(* IEC 61131-3 sources: STruCpp/libs/sources/plcopen-softmotion, 17 files *)

(* ---- opensml_axis.st ---- *)
(*
 * OpenSML_Axis — CiA 402 axis reference structure.
 *
 * Vendored from OpenSML (https://github.com/feecat/OpenSML), GPL-3.0.
 * Each field maps 1:1 onto a CiA 402 drive object exchanged over the
 * fieldbus (e.g. EtherCAT PDOs). Outputs (%Q) are written by the motion
 * blocks; inputs (%I) are read from the drive each scan.
 *)
TYPE OpenSML_Axis :
STRUCT
	(* Outputs -> drive *)
	ControlWord : UINT;                 (* 0x6040 *)
	Modes_of_operation : SINT;          (* 0x6060 *)
	Target_Position : DINT;             (* 0x607A *)
	Profile_Velocity : UDINT;           (* 0x6081 *)
	Target_Velocity : DINT;             (* 0x60FF *)
	Target_torque : INT;                (* 0x6071 *)
	(* Inputs <- drive *)
	StatusWord : UINT;                  (* 0x6041 *)
	Modes_of_operation_display : SINT;  (* 0x6061 *)
	Torque_Actual_Value : INT;          (* 0x6077 *)
	Position_Actual_Value : DINT;       (* 0x6064 *)
	Velocity_Actual_Value : DINT;       (* 0x606C *)
	Current_Actual_Value : INT;         (* 0x6078 *)
	Following_Error_Actual_Value : DINT;(* 0x60F4 *)
END_STRUCT
END_TYPE

(* ---- opensml_control.st ---- *)
(*
 * OpenSML_Control — aggregate axis command/status structure.
 * Vendored from OpenSML (https://github.com/feecat/OpenSML), GPL-3.0.
 *)
TYPE OpenSML_Control :
STRUCT
	xAxisEnable: BOOL;//Axis Hardware Enable
	xMoveEnable: BOOL;//Jog&Pos Movement Enable
	xHomeEnable: BOOL;//Home Function Enable
	xSimulation: BOOL;//Simulation Mode
	xEmergencyStop: BOOL:=TRUE;//Emergency Stop

	JogPos: BOOL;//Jog Positive
	JogNeg: BOOL;//Jog Negative
	JogVelocity: LREAL:=10;//Jog Velocity

	lrActualPosition: LREAL;//Actual Position Feedback

	lrFollowPosition: LREAL;//Follow Target Position, Can be set to new value at any time
	lrFollowVelocity: LREAL:=20;//Follow Move Velocity, Can be set to new value at any time
	xFollowEnable: BOOL;//Follow Move Enable

	xError: BOOL;//Error
	xBusy: BOOL;//Busy, Normal Working State
	xInPosition: BOOL;//In Position
	xEnabled: BOOL;//Axis Hardware Enabled
	xHomeDone: BOOL;//Axis Home Done

	MaxVelocity: LREAL:=100;//Max Velocity
	MaxAcceleration: LREAL:=1000;//Max Acceleration
	MaxJerk: LREAL:=10000;//Max Jerk
	CycleTime: LREAL:=0.001;//Task Cycle Time, 0.001 = 1ms
	Scale: LREAL:=16#1000;//Scale

	Axis:OpenSML_Axis;//Axis Reference
END_STRUCT
END_TYPE

(* ---- s7rtt_types.st ---- *)
(*
 * S7RTT motion-state / limits structures.
 * Vendored from S7RTT (https://github.com/feecat/S7RTT), Apache-2.0.
 * Converted from PLCopen XML. Single-axis 7-segment S-curve OTG.
 *)

TYPE ST_MotionLimits :
STRUCT
	fVelMax : LREAL;
	fAccMax : LREAL;
	fJerkMax : LREAL;
END_STRUCT
END_TYPE

TYPE ST_MotionState :
STRUCT
	fDuration : LREAL := 0.0;
	fPos : LREAL := 0.0;
	fVel : LREAL := 0.0;
	fAcc : LREAL := 0.0;
	fJerk : LREAL := 0.0;
END_STRUCT
END_TYPE

(* ---- sm3_axis_ref.st ---- *)
(*
 * AXIS_REF_SM3 — CODESYS SoftMotion-compatible axis reference.
 *
 * Application code declares an axis of this type (the EtherCAT drive's name),
 * passes it to MC_* blocks by VAR_IN_OUT, and reads/writes its fields
 * (fActPosition, nAxisState, …) — exactly as in CODESYS. It is a STRUCT (not an
 * FB): real CODESYS application code never calls axis methods (those are all
 * driver-internal). All positions/velocities are in technical (user) units;
 * the embedded `Drive` carries the raw CiA 402 PDO words in increments, and
 * SM_Drive_GenericDS402 bridges between them each scan.
 *)
TYPE AXIS_REF_SM3 :
STRUCT
	(* --- Command (written by MC_* blocks, in technical units) --- *)
	fSetPosition : LREAL;              (* commanded position [u] *)
	fSetVelocity : LREAL;              (* commanded velocity [u/s] *)
	fSetAcceleration : LREAL;          (* commanded acceleration [u/s2] *)
	fSetDeceleration : LREAL;          (* commanded deceleration [u/s2] *)
	fSetJerk : LREAL;                  (* commanded jerk [u/s3] *)
	bRegulatorOn : BOOL;               (* power-stage enable command *)
	bDriveStart : BOOL;                (* quick-stop release command *)
	byControllerMode : BYTE;           (* SMC_CONTROLLER_MODE as BYTE *)

	(* --- Feedback (updated by the drive bridge, in technical units) --- *)
	fActPosition : LREAL;              (* actual position [u] *)
	fActVelocity : LREAL;              (* actual velocity [u/s] *)
	fActTorque : LREAL;                (* actual torque *)
	nAxisState : SMC_AXIS_STATE;       (* PLCopen axis state *)
	bRegulatorRealState : BOOL;        (* real power-stage state *)
	bDriveStartRealState : BOOL;       (* real quick-stop-released state *)
	byRealControllerMode : BYTE;       (* actual controller mode *)

	(* --- Error / communication --- *)
	bError : BOOL;
	dwErrorID : DWORD;                 (* SMC_ERROR as DWORD *)
	bCommunication : BOOL;
	wCommunicationState : WORD;

	(* --- Scaling (increments <-> technical units) --- *)
	iRatioTechUnitsNum : DINT := 1;    (* CODESYS param 1052 *)
	dwRatioTechUnitsDenom : DWORD := 1;(* CODESYS param 1051 *)
	fScalefactor : LREAL := 1.0;       (* CODESYS param 1054 *)
	fIncPerUnit : LREAL := 1.0;        (* derived: increments per user unit *)

	(* --- Axis configuration --- *)
	fPositionPeriod : LREAL := 360.0;  (* modulo period [u] *)
	bModulo : BOOL;                    (* TRUE = rotary/modulo axis *)
	fSWLimitPositive : LREAL;
	fSWLimitNegative : LREAL;
	bSWLimitEnable : BOOL;
	fCycleTime : LREAL := 0.01;        (* task cycle [s], for OTG *)

	(* --- Raw CiA 402 interface (increments) bridged to the drive PDOs --- *)
	Drive : OpenSML_Axis;
END_STRUCT
END_TYPE

(* ---- sm3_enums.st ---- *)
(*
 * CODESYS SoftMotion (SM3) compatible enum types.
 *
 * Values follow CODESYS SM3_Basic / SM3_Error so that ported application code
 * comparing against these names/values behaves identically. This is the
 * single-axis CiA 402 subset (see docs/PLCOPEN_SOFTMOTION_ETHERCAT_PLAN.md).
 *)

(* PLCopen axis state (AXIS_REF_SM3.nAxisState) *)
TYPE SMC_AXIS_STATE : (
	power_off := 0,
	errorstop := 1,
	stopping := 2,
	standstill := 3,
	discrete_motion := 4,
	continuous_motion := 5,
	synchronized_motion := 6,
	homing := 7
); END_TYPE

(* Controller mode (AXIS_REF_SM3.byControllerMode / SMC_SetControllerMode) *)
TYPE SMC_CONTROLLER_MODE : (
	SMC_nocontrol := 0,
	SMC_torque := 1,
	SMC_velocity := 2,
	SMC_position := 3,
	SMC_current := 4
); END_TYPE

(* Movement direction for MC_MoveAbsolute / MC_MoveVelocity (modulo axes) *)
TYPE MC_DIRECTION : (
	mcd_negative := -1,
	mcd_current := 0,
	mcd_positive := 1,
	mcd_shortest := 2,
	mcd_fastest := 3
); END_TYPE

(* Buffering behaviour relative to a preceding motion command *)
TYPE MC_BUFFER_MODE : (
	mcbm_aborting := 0,
	mcbm_buffered := 1,
	mcbm_blending_low := 2,
	mcbm_blending_previous := 3,
	mcbm_blending_next := 4,
	mcbm_blending_high := 5
); END_TYPE

(* Homing mode (subset — the CiA 402 relevant ones) *)
TYPE SMC_HOMING_MODE : (
	smc_hm_direct := 0,
	smc_hm_limit_switch := 1,
	smc_hm_reference_pulse := 2,
	smc_hm_drive_internal := 35
); END_TYPE

(*
 * Error identifier (MC_*.ErrorID). Single-axis CiA 402 subset of CODESYS
 * SMC_ERROR (the 0..~500 drive-interface / limits / controller-mode /
 * FB-input band). Values match CODESYS where documented.
 *)
TYPE SMC_ERROR : (
	SMC_NO_ERROR := 0,
	SMC_DI_GENERAL_COMMUNICATION_ERROR := 1,
	SMC_DI_AXIS_ERROR := 2,
	SMC_DI_SWLIMITS_EXCEEDED := 10,
	SMC_DI_HWLIMITS_EXCEEDED := 11,
	SMC_DI_HALT_OR_QUICKSTOP_NOT_SUPPORTED := 12,
	SMC_DI_VOLTAGE_DISABLED := 13,
	SMC_DI_FIELDBUS_LOST_SYNCRONITY := 14,
	SMC_DI_COMMUNICATION_INTERRUPTED := 15,
	SMC_REGULATOR_OR_START_NOT_SET := 20,
	SMC_WRONG_CONTROLLER_MODE := 21,
	SMC_FB_WASNT_CALLED_DURING_MOTION := 22,
	SMC_AXIS_IS_NO_AXIS_REF := 23,
	SMC_AXIS_REF_CHANGED_DURING_OPERATION := 24,
	SMC_FB_ACTIVE_AXIS_DISABLED := 25,
	SMC_AXIS_NOT_READY_FOR_MOTION := 26,
	SMC_NicNyet_ERROR := 30,
	SMC_MA_INVALID_ACCDEC_VALUES := 110,
	SMC_MA_INVALID_DIRECTION := 111,
	SMC_MV_INVALID_VELACC_VALUES := 120,
	SMC_MV_DIRECTION_NOT_APPLICABLE := 121,
	SMC_H_AXIS_WASNT_STANDING_STILL := 130,
	SMC_H_AXIS_DIDNT_START_HOMING := 131,
	SMC_H_HOMING_TIMEOUT := 132,
	SMC_R_NO_ERROR_TO_RESET := 140,
	SMC_R_DRIVE_DOESNT_ANSWER := 141,
	SMC_STOP_ERROR_DURING_STOP := 150,
	SMC_3SH_INVALID_VELACC_VALUES := 160
); END_TYPE

(* ---- s7rtt_functions.st ---- *)
(*
 * S7RTT trajectory helper functions (AtTime / BuildProfile / CalcTrajDist).
 * Vendored from S7RTT (https://github.com/feecat/S7RTT), Apache-2.0.
 * Converted from PLCopen XML. Single-axis 7-segment S-curve OTG.
 *)

FUNCTION FC_S7RTT_AtTime : ST_MotionState
VAR_INPUT
	Trajectory : ARRAY[1..32] OF ST_MotionState;
	SegCount : INT;
	ElapsedTime : LREAL;
END_VAR
VAR
	i : INT;
	t_rem : LREAL;
	t : LREAL;
	j : LREAL;
	p0 : LREAL;
	v0 : LREAL;
	a0 : LREAL;
	last_idx : INT;
END_VAR

IF SegCount <= 0 THEN
    // No trajectory, return first state
    FC_S7RTT_AtTime.fPos := Trajectory[1].fPos; FC_S7RTT_AtTime.fVel := 0.0; FC_S7RTT_AtTime.fAcc := 0.0;
    RETURN;
END_IF;

IF ElapsedTime <= 0.0 THEN
     // Return Initial State from First Segment
     FC_S7RTT_AtTime := Trajectory[1];
     FC_S7RTT_AtTime.fDuration := 0.0;
     FC_S7RTT_AtTime.fJerk := 0.0;
     RETURN;
END_IF;

t_rem := ElapsedTime;

FOR i := 1 TO SegCount DO
	IF t_rem <= Trajectory[i].fDuration THEN
		t := t_rem;
		j := Trajectory[i].fJerk;
		// Use pre-calculated state at segment start
		p0 := Trajectory[i].fPos;
		v0 := Trajectory[i].fVel;
		a0 := Trajectory[i].fAcc;

		FC_S7RTT_AtTime.fPos := p0 + v0 * t + 0.5 * a0 * t*t + (1.0/6.0) * j * t*t*t;
		FC_S7RTT_AtTime.fVel := v0 + a0 * t + 0.5 * j * t*t;
		FC_S7RTT_AtTime.fAcc := a0 + j * t;
		FC_S7RTT_AtTime.fJerk := j;
		FC_S7RTT_AtTime.fDuration := 0.0;
		RETURN;
	ELSE
		t_rem := t_rem - Trajectory[i].fDuration;
	END_IF;
END_FOR;

// Time is beyond end of trajectory
// Calculate Final State of last segment
last_idx := SegCount;
t := Trajectory[last_idx].fDuration;
j := Trajectory[last_idx].fJerk;
p0 := Trajectory[last_idx].fPos;
v0 := Trajectory[last_idx].fVel;
a0 := Trajectory[last_idx].fAcc;

p0 := p0 + v0 * t + 0.5 * a0 * t*t + (1.0/6.0) * j * t*t*t;
v0 := v0 + a0 * t + 0.5 * j * t*t;

// Hold Final Position (assuming v=target, a=0 at end)
// Linear projection if Velocity is non-zero
FC_S7RTT_AtTime.fPos := p0 + v0 * t_rem;
FC_S7RTT_AtTime.fVel := v0;
FC_S7RTT_AtTime.fAcc := 0.0;
FC_S7RTT_AtTime.fJerk := 0.0;
FC_S7RTT_AtTime.fDuration := 0.0;
END_FUNCTION

FUNCTION FC_S7RTT_BuildProfile : INT
VAR_INPUT
	in_v_start : LREAL;
	in_a_start : LREAL;
	in_v_target : LREAL;
	in_a_max : LREAL;
	in_j_max : LREAL;
END_VAR
VAR_IN_OUT
	out_time : ARRAY[1..5] OF LREAL;
	out_jerk : ARRAY[1..5] OF LREAL;
END_VAR
VAR
	acc_clamped : LREAL;
	t_to_zero : LREAL;
	j_restore : LREAL;
	v_min_feasible : LREAL;
	direction : LREAL;
	v0_mod : LREAL;
	a0_mod : LREAL;
	v1_mod : LREAL;
	t1_max : LREAL;
	t3_max : LREAL;
	dv_inflection : LREAL;
	dv_req : LREAL;
	dv_missing : LREAL;
	term : LREAL;
	a_peak : LREAL;
	t1 : LREAL;
	t2 : LREAL;
	t3 : LREAL;
	cnt : INT;
	EPS : LREAL := 1E-10;
END_VAR

cnt := 0;

// 1. Clamp initial acceleration to limits
acc_clamped := in_a_start;
IF acc_clamped > in_a_max THEN acc_clamped := in_a_max; END_IF;
IF acc_clamped < -in_a_max THEN acc_clamped := -in_a_max; END_IF;

// 2. Check feasibility (can we stop?)
t_to_zero := ABS(acc_clamped) / in_j_max;
IF ABS(acc_clamped) > EPS THEN
    IF acc_clamped > 0.0 THEN j_restore := -in_j_max; ELSE j_restore := in_j_max; END_IF;
ELSE
    j_restore := 0.0;
END_IF;

v_min_feasible := in_v_start + acc_clamped * t_to_zero + 0.5 * j_restore * t_to_zero * t_to_zero;

// 3. Determine direction
direction := 1.0;
IF in_v_target < v_min_feasible - EPS THEN
    direction := -1.0;
END_IF;

// 4. Normalize to positive quadrant
v0_mod := in_v_start * direction;
a0_mod := acc_clamped * direction;
v1_mod := in_v_target * direction;

t1_max := (in_a_max - a0_mod) / in_j_max;
IF t1_max < 0.0 THEN t1_max := 0.0; END_IF;

t3_max := in_a_max / in_j_max;

// Velocity change at inflection (max accel reached)
dv_inflection := (a0_mod * t1_max + 0.5 * in_j_max * t1_max * t1_max) +
                 (in_a_max * t3_max - 0.5 * in_j_max * t3_max * t3_max);

dv_req := v1_mod - v0_mod;

// 5. Calculate profile times
IF dv_req > dv_inflection THEN
    // Trapezoidal (Constant Acceleration Phase)
    dv_missing := dv_req - dv_inflection;
    t2 := dv_missing / in_a_max;
    t1 := t1_max;
    t3 := t3_max;
ELSE
    // Triangular (No Constant Acceleration)
    term := in_j_max * dv_req + 0.5 * a0_mod * a0_mod;
    IF term < 0.0 THEN term := 0.0; END_IF;
    a_peak := SQRT(term);

    t1 := (a_peak - a0_mod) / in_j_max;
    IF t1 < 0.0 THEN t1 := 0.0; END_IF;

    t3 := a_peak / in_j_max;
    IF t3 < 0.0 THEN t3 := 0.0; END_IF;

    t2 := 0.0;
END_IF;

// 6. Output Segments
IF t1 > EPS THEN
    cnt := cnt + 1; out_time[cnt] := t1; out_jerk[cnt] := direction * in_j_max;
END_IF;
IF t2 > EPS THEN
    cnt := cnt + 1; out_time[cnt] := t2; out_jerk[cnt] := 0.0;
END_IF;
IF t3 > EPS THEN
    cnt := cnt + 1; out_time[cnt] := t3; out_jerk[cnt] := -direction * in_j_max;
END_IF;

FC_S7RTT_BuildProfile := cnt;
END_FUNCTION

FUNCTION FC_S7RTT_CalcTrajDist : LREAL
VAR_INPUT
	v_peak : LREAL;
	start_v : LREAL;
	start_a : LREAL;
	target_v : LREAL;
	a_max : LREAL;
	j_max : LREAL;
END_VAR
VAR
	t_buf : ARRAY[1..5] OF LREAL;
	j_buf : ARRAY[1..5] OF LREAL;
	cnt : INT;
	i : INT;
	v_curr : LREAL;
	a_curr : LREAL;
	dist_total : LREAL;
	t_seg : LREAL;
	j_seg : LREAL;
END_VAR

dist_total := 0.0;
v_curr := start_v;
a_curr := start_a;

// Phase 1: Start -> Peak Velocity
cnt := FC_S7RTT_BuildProfile(v_curr, a_curr, v_peak, a_max, j_max, t_buf, j_buf);
FOR i := 1 TO cnt DO
	t_seg := t_buf[i];
	j_seg := j_buf[i];
    // Standard kinematic integration: p = p0 + v0*t + 0.5*a0*t^2 + 1/6*j*t^3
	dist_total := dist_total + v_curr * t_seg + 0.5 * a_curr * t_seg*t_seg + (1.0/6.0) * j_seg * t_seg*t_seg*t_seg;
	v_curr := v_curr + a_curr * t_seg + 0.5 * j_seg * t_seg*t_seg;
	a_curr := a_curr + j_seg * t_seg;
END_FOR;

// Phase 2: Peak Velocity -> Target Velocity
cnt := FC_S7RTT_BuildProfile(v_curr, a_curr, target_v, a_max, j_max, t_buf, j_buf);
FOR i := 1 TO cnt DO
	t_seg := t_buf[i];
	j_seg := j_buf[i];
	dist_total := dist_total + v_curr * t_seg + 0.5 * a_curr * t_seg*t_seg + (1.0/6.0) * j_seg * t_seg*t_seg*t_seg;
	v_curr := v_curr + a_curr * t_seg + 0.5 * j_seg * t_seg*t_seg;
	a_curr := a_curr + j_seg * t_seg;
END_FOR;

FC_S7RTT_CalcTrajDist := dist_total;
END_FUNCTION

(* ---- opensml_axis_controller.st ---- *)
(*
 * OpenSML_AxisController — high-level jog/follow controller over OpenSML_Control.
 * Vendored from OpenSML (https://github.com/feecat/OpenSML), GPL-3.0.
 *)
FUNCTION_BLOCK OpenSML_AxisController
VAR_IN_OUT
	Axis:OpenSML_Axis;
	Control:OpenSML_Control;
END_VAR
VAR
	Power:OpenSML_Power;
	Home:OpenSML_Home;
	iState:INT;
	otg : FB_S7RTT_OTG;
	InterfaceType:BOOL;
	JogVel:LREAL;
	MoveVel:LREAL;
END_VAR

Power(
	Axis:=Axis ,
	xEnable:=Control.xAxisEnable ,
	xEmergencyStop:=Control.xEmergencyStop ,
	xDone=>Control.xEnabled );

Home(
	Axis:=Axis ,
	xEnable:=Control.xHomeEnable AND NOT Control.xMoveEnable ,
	xDone=>Control.xHomeDone );

(*
Cyclic Synchronous Position Mode (=8)
Set 6060(Op mode) and 60C2(Interpolation time period) at Startup Parameters.

#####################################
NEED StruckigLight Library for Quadratic Velocity Ramp Calculate.

If in movement, Please DO NOT Drop down xEnable.
#####################################
*)

Control.xInPosition:=FALSE;

IF control.xSimulation THEN
	Axis.Position_Actual_Value:=Axis.Target_Position;
END_IF

control.lrActualPosition:=DINT_TO_LREAL(Axis.Position_Actual_Value) / Control.Scale;

CASE iState OF
	0://start
		Control.xError:=FALSE;
		IF Control.xMoveEnable AND Axis.StatusWord.1 AND Axis.StatusWord.2 AND Axis.Modes_of_operation_display = 8 AND NOT Axis.StatusWord.3 THEN//ready
			iState:=10;//go go
		ELSIF Control.xMoveEnable AND Axis.StatusWord.1 AND Axis.Modes_of_operation_display <> 8 THEN//need switch mode
			Axis.ControlWord.3:=FALSE;//drop down operation enabled, motor could free move
			iState:=10;
		ELSIF Control.xMoveEnable AND Control.xSimulation THEN
			iState:=20;
		ELSIF Control.xMoveEnable THEN
			iState:=999;//error
		END_IF
	10://Set Mode
		Axis.Modes_of_operation:=8;//Cyclic Synchronous Position Mode
		Axis.ControlWord.3:=Axis.Modes_of_operation_display=8;//Success change mode, enable operation
		otg.CurrentPosition:=DINT_TO_LREAL(Axis.Position_Actual_Value) / Control.Scale;//Write actual position to otg
		IF Axis.StatusWord.2 AND Axis.Modes_of_operation_display = 8 THEN//Operation Enabled, Mode Changed success
			iState:=20;
		END_IF
	20://Movement
		IF Control.JogPos AND NOT Control.xFollowEnable THEN
			InterfaceType:=1;
			JogVel:=MIN(Control.JogVelocity, Control.MaxVelocity);
		ELSIF Control.JogNeg AND NOT Control.xFollowEnable THEN
			InterfaceType:=1;
			JogVel:=MAX(-Control.JogVelocity, -Control.MaxVelocity);
		ELSE
			InterfaceType:=1;
			JogVel:=0;
		END_IF

		IF Control.xFollowEnable AND Control.lrFollowVelocity > 0 THEN
			InterfaceType:=0;
			MoveVel:=MIN(Control.lrFollowVelocity, Control.MaxVelocity);
		ELSE
			MoveVel:= Control.MaxVelocity;
		END_IF

		otg(
			ControlInterface:= InterfaceType,
			TargetPosition:= Control.lrFollowPosition ,
			TargetVelocity:= JogVel ,
			CycleTIme:= Control.CycleTime,
			MaxVelocity:= MoveVel,//Control.para.MaxVelocity ,
			MaxAcceleration:= Control.MaxAcceleration ,
			MaxJerk:= Control.MaxJerk);//accept new position and going on

		IF otg.NewPosition >= 0 THEN
			Axis.Target_Position := LREAL_TO_DINT(otg.NewPosition * Control.Scale);
		ELSE
			Axis.Target_Position := - LREAL_TO_DINT( - otg.NewPosition * Control.Scale);//it fix negative overflow problem.
		END_IF

		Control.xInPosition := ABS(otg.NewPosition - Control.lrActualPosition) < 0.01;

		IF Axis.StatusWord.13 OR Axis.StatusWord.3 OR otg.xError OR Power.xError OR Home.xError THEN//Axis Error
			iState:=999;
		ELSIF NOT Control.xMoveEnable THEN
			iState:=0;
		END_IF
	999://Error wait
		Control.xError:=TRUE;
		IF NOT Control.xMoveEnable THEN
			iState:=0;
		END_IF
END_CASE

END_FUNCTION_BLOCK

(* ---- opensml_home.st ---- *)
(*
 * Homing (CiA402 mode 6)
 * Vendored from OpenSML (https://github.com/feecat/OpenSML), GPL-3.0.
 * Part of the strucpp plcopen-softmotion bundled library.
 *)
FUNCTION_BLOCK OpenSML_Home
VAR_IN_OUT
	Axis:OpenSML_Axis;
END_VAR
VAR_INPUT
	xEnable:BOOL;
END_VAR
VAR_OUTPUT
	xDone:BOOL;
	xError:BOOL;
END_VAR
VAR
	iState:INT;
	tonTimeout:TON;
	Pos_Old:DINT;
END_VAR

(*
Home Function Block
Need Manually Write To SDO:
607C: Home Offset
6098: Home method
6099: Home Speeds*
609A: Home Acceleration

6099.01 - Home Speed for Search Limit Switch
6099.02 - Home Speed for Index Pulse
*)
CASE iState OF
	0:
		xDone:=FALSE;
		xError:=FALSE;
		IF xEnable AND Axis.StatusWord.1 AND Axis.StatusWord.2 AND Axis.Modes_of_operation_display = 6 AND NOT Axis.StatusWord.3 THEN//ready
			iState:=10;//go go
		ELSIF xEnable AND Axis.StatusWord.1 AND Axis.Modes_of_operation_display <> 6 THEN//need switch mode
			Axis.ControlWord.3:=FALSE;//drop down operation enabled
			iState:=10;
		ELSIF xEnable THEN
			iState:=999;//error
		END_IF
	10:
		Axis.ControlWord.4 := FALSE;//Reset reference bit
		Axis.Modes_of_operation:=6;//Home Mode
		Axis.ControlWord.3:=Axis.Modes_of_operation_display=6;//Success change mode, enable operation
		IF Axis.StatusWord.2 THEN//Operation Enabled
			iState:=20;
		END_IF
	20:
		Axis.ControlWord.4 := TRUE;//start reference
		tonTimeout(IN:=axis.Position_Actual_Value = Pos_Old, pt:=T#10S);//If Position didnt change, error
		Pos_Old:=Axis.Position_Actual_Value;
		IF Axis.StatusWord.12 THEN//If HomeAttained, Success
			tonTimeout(IN:=FALSE);
			Axis.ControlWord.4:=FALSE;
			Axis.Target_Position:=Axis.Position_Actual_Value;
			iState:=30;
		ELSIF tonTimeout.Q OR NOT xEnable OR Axis.StatusWord.3 OR Axis.StatusWord.13 THEN iState:=999;//error
		END_IF
	30:
		xDone:=TRUE;
		IF NOT xEnable THEN//Wait next home
			iState:=0;
		END_IF
	999:
		tonTimeout(IN:=FALSE);
		Axis.ControlWord.4:=FALSE;
		xError:=TRUE;
		IF NOT xEnable THEN
			iState:=0;
		END_IF
END_CASE

END_FUNCTION_BLOCK

(* ---- opensml_power.st ---- *)
(*
 * MC_Power power stage / CiA402 enable sequence
 * Vendored from OpenSML (https://github.com/feecat/OpenSML), GPL-3.0.
 * Part of the strucpp plcopen-softmotion bundled library.
 *)
FUNCTION_BLOCK OpenSML_Power
VAR_IN_OUT
	Axis:OpenSML_Axis;
END_VAR
VAR_INPUT
	xEnable: BOOL;
	xEmergencyStop: BOOL:=TRUE;
END_VAR
VAR_OUTPUT
	xDone: BOOL;
	xError: BOOL;
END_VAR
VAR
	iState:INT;
	tonTimeout:TON;
	tTimeOut:TIME:=T#500MS;
END_VAR

(*
MC_Power
Can Also be used MC_Reset, just trigger xEnable.
It is Highly Recommend to use OpenSML_Stop to force stop movements.
*)
Axis.ControlWord.2:=xEmergencyStop;//QuickStop
CASE iState OF
	0://start
		xDone:=FALSE;
		xError:=FALSE;
		Axis.ControlWord.0:=FALSE;//SwitchOn
		Axis.ControlWord.1:=FALSE;//EnableVoltage
		Axis.ControlWord.3:=FALSE;//EnableOperation
		Axis.ControlWord.7:=FALSE;//FaultReset
		IF xEnable THEN
			IF Axis.StatusWord.3 THEN iState:=10;//If there have error, Reset first
			ELSE iState:=20;//No error, go go
			END_IF
		END_IF
	10://reset
		Axis.ControlWord.7:=TRUE;//bit7 faultreset
		tonTimeout(IN:=TRUE,PT:=tTimeOut);
		IF tonTimeout.Q AND NOT Axis.StatusWord.3 THEN//not fault
			Axis.ControlWord.7:=FALSE;//bit7 faultreset
			tonTimeout(IN:=FALSE);
			iState:=20;
		ELSIF tonTimeout.Q THEN iState:=999;//error
		END_IF
	20://Enable Voltage
		Axis.ControlWord.1:=TRUE;
		tonTimeout(IN:=TRUE,PT:=tTimeOut);
		IF Axis.StatusWord.0 THEN//ReadyToSwitchOn
			tonTimeout(IN:=FALSE);
			iState:=30;
		ELSIF tonTimeout.Q THEN iState:=999;//error
		END_IF
	30://Switch ON
		Axis.ControlWord.0:=TRUE;
		tonTimeout(IN:=TRUE,pt:=tTimeOut);
		IF Axis.StatusWord.1 THEN
			tonTimeout(IN:=FALSE);
			iState:=40;
		ELSIF tonTimeout.Q THEN iState:=999;//error
		END_IF
	40://EnableOperation
		Axis.Target_Position:=Axis.Position_Actual_Value;
		Axis.ControlWord.3:=TRUE;
		tonTimeout(IN:=TRUE,pt:=tTimeOut);
		IF Axis.StatusWord.2 THEN
			tonTimeout(IN:=FALSE);
			iState:=50;
		ELSIF tonTimeout.Q THEN iState:=999;//error
		END_IF
	50://Success
		xDone:=TRUE;
		IF NOT xEnable THEN
			Axis.ControlWord.3:=FALSE;
			iState:=0;
		END_IF
		IF Axis.StatusWord.3 THEN
			iState:=999;//Error when running
		END_IF
	999://Error wait
		tonTimeout(IN:=FALSE);
		xError:=TRUE;
		IF NOT xEnable THEN
			iState:=0;
		END_IF
END_CASE

END_FUNCTION_BLOCK

(* ---- opensml_profile_position.st ---- *)
(*
 * Profile Position mode (CiA402 mode 1)
 * Vendored from OpenSML (https://github.com/feecat/OpenSML), GPL-3.0.
 * Part of the strucpp plcopen-softmotion bundled library.
 *)
FUNCTION_BLOCK OpenSML_ProfilePosition
VAR_IN_OUT
	Axis:OpenSML_Axis;
END_VAR
VAR_INPUT
	xEnable:BOOL;
	xExecute: BOOL;
	xContinueMove: BOOL;
	xRelativeMode: BOOL;
	diTargetPosition:DINT;
	udiProfileVelocity:UDINT;
END_VAR
VAR_OUTPUT
	xDone: BOOL;
	xBusy: BOOL;
	xMoving: BOOL;
	xError: BOOL;
END_VAR
VAR
	iState:INT;
	tonTimeout:TON;
	tTimeOut:TIME:=T#200MS;
END_VAR

(*
Profile Position Mode (=1)
Manually Write To SDO or Write To PDO If Needed:
6083: Profile Acceleration
6084: Profile Deceleration
6085: Quick Stop Deceleration
*)
//Settings
Axis.ControlWord.5:=xContinueMove;//It means if 1st positon not arrived and there got 2st position, It Will No Deceleration And continues the movements.
Axis.ControlWord.6:=xRelativeMode;//0 is Absolute, 1 is Relative
Axis.ControlWord.4:=xExecute AND iState = 20;
xBusy:=iState=20 AND Axis.StatusWord.12 AND NOT Axis.StatusWord.10;//Acknowledge and not Reached
xDone:=iState=20 AND Axis.StatusWord.10 AND NOT Axis.StatusWord.13;//Target Reached and not Following Error
xMoving:=NOT Axis.StatusWord.14;//Not Standstill

CASE iState OF
	0://start
		xDone:=FALSE;
		xBusy:=FALSE;
		xError:=FALSE;
		IF xEnable AND Axis.StatusWord.1 AND Axis.StatusWord.2 AND Axis.Modes_of_operation_display = 1 AND NOT Axis.StatusWord.3 THEN//ready
			iState:=10;//go go
		ELSIF xEnable AND Axis.StatusWord.1 AND Axis.Modes_of_operation_display <> 1 THEN//need switch mode
			Axis.ControlWord.3:=FALSE;//drop down operation enabled
			iState:=10;
		ELSIF xEnable THEN
			iState:=999;//error
		END_IF
	10://Set Mode
		Axis.Modes_of_operation:=1;//Profile Position Mode
		Axis.ControlWord.3:=Axis.Modes_of_operation_display=1;//Success change mode, enable operation
		IF Axis.StatusWord.2 AND Axis.Modes_of_operation_display = 1 THEN//Operation Enabled, Mode Changed success
			iState:=20;
		END_IF
	20://Movement
		Axis.Profile_Velocity:=udiProfileVelocity;
		Axis.Target_Position:=diTargetPosition;
		IF Axis.StatusWord.13 OR Axis.StatusWord.3 THEN//Axis Error
			iState:=999;
		ELSIF NOT xEnable THEN
			Axis.Profile_Velocity:=0;
			Axis.Target_Position:=0;
			iState:=0;
		END_IF
	999://Error wait
		Axis.Profile_Velocity:=0;
		Axis.Target_Position:=0;
		tonTimeout(IN:=FALSE);
		xError:=TRUE;
		IF NOT xEnable THEN
			iState:=0;
		END_IF
END_CASE

END_FUNCTION_BLOCK

(* ---- opensml_profile_velocity.st ---- *)
(*
 * Profile Velocity mode (CiA402 mode 3)
 * Vendored from OpenSML (https://github.com/feecat/OpenSML), GPL-3.0.
 * Part of the strucpp plcopen-softmotion bundled library.
 *)
FUNCTION_BLOCK OpenSML_ProfileVelocity
VAR_IN_OUT
	Axis:OpenSML_Axis;
END_VAR
VAR_INPUT
	xEnable:BOOL;
	diTargetVelocity:DINT;
END_VAR
VAR_OUTPUT
	xError: BOOL;
END_VAR
VAR
	iState:INT;
	tonTimeout:TON;
	tTimeOut:TIME:=T#200MS;
END_VAR

(*
Profile Velocity Mode (=3)
Manually Write To SDO or Write To PDO If Needed:
6083: Profile Acceleration
6084: Profile Deceleration
6085: Quick Stop Deceleration
*)
CASE iState OF
	0://start
		xError:=FALSE;
		IF xEnable AND Axis.StatusWord.1 AND Axis.StatusWord.2 AND Axis.Modes_of_operation_display = 3 AND NOT Axis.StatusWord.3 THEN//ready
			iState:=10;//go go
		ELSIF xEnable AND Axis.StatusWord.1 AND Axis.Modes_of_operation_display <> 3 THEN//need switch mode
			Axis.ControlWord.3:=FALSE;//drop down operation enabled
			iState:=10;
		ELSIF xEnable THEN
			iState:=999;//error
		END_IF
	10://Set Mode
		Axis.Modes_of_operation:=3;//Profile Velocity Mode
		Axis.ControlWord.3:=Axis.Modes_of_operation_display=3;//Success change mode, enable operation
		IF Axis.StatusWord.2 AND Axis.Modes_of_operation_display = 3 THEN//Operation Enabled, Mode Changed success
			iState:=20;
		END_IF
	20://Movement
		Axis.Target_Velocity:=diTargetVelocity;
		IF Axis.StatusWord.3 THEN
			iState:=999;
		ELSIF NOT xEnable THEN
			Axis.Target_Velocity:=0;
			iState:=0;
		END_IF
	999://Error wait
		Axis.Target_Velocity:=0;
		tonTimeout(IN:=FALSE);
		xError:=TRUE;
		IF NOT xEnable THEN
			iState:=0;
		END_IF
END_CASE

END_FUNCTION_BLOCK

(* ---- opensml_stop.st ---- *)
(*
 * Software stop (halt bit)
 * Vendored from OpenSML (https://github.com/feecat/OpenSML), GPL-3.0.
 * Part of the strucpp plcopen-softmotion bundled library.
 *)
FUNCTION_BLOCK OpenSML_Stop
VAR_IN_OUT
	Axis:OpenSML_Axis;
END_VAR
VAR_INPUT
	xStop: BOOL;
END_VAR
VAR_OUTPUT
END_VAR
VAR
END_VAR

(*
MC_Stop
Software Stop, True=Stop
*)
Axis.ControlWord.8:=xStop;
END_FUNCTION_BLOCK

(* ---- opensml_sync_position.st ---- *)
(*
 * OpenSML Cyclic Synchronous Position (CiA402 mode 8) via S7RTT OTG.
 * Vendored from OpenSML (https://github.com/feecat/OpenSML), GPL-3.0.
 *)
FUNCTION_BLOCK OpenSML_SyncPosition
VAR_IN_OUT
	Axis:OpenSML_Axis;
END_VAR
VAR_INPUT
	MaxVelocity :LREAL:=2000;
	MaxAcceleration :LREAL:=200;
	MaxJerk :LREAL:=200;
	CycleTime:LREAL:=0.001;//0.001 = 1ms

	TargetPosition :LREAL;
	xEnable: BOOL;
	lrScale:LREAL:=1.0;
	xSimulation: BOOL;	// added: referenced in body but undeclared upstream
END_VAR
VAR_OUTPUT
	xError: BOOL;
END_VAR
VAR
	otg : FB_S7RTT_OTG;
	iState:INT;

END_VAR

(*
Cyclic Synchronous Position Mode (=8)
Set 6060(Op mode) and 60C2(Interpolation time period) at Startup Parameters.

#####################################
NEED StruckigLight Library for Quadratic Velocity Ramp Calculate.

If in movement, Please DO NOT Drop down xEnable.
#####################################
*)

CASE iState OF
	0://start
		xError:=FALSE;
		IF xEnable AND Axis.StatusWord.1 AND Axis.StatusWord.2 AND Axis.Modes_of_operation_display = 8 AND NOT Axis.StatusWord.3 THEN//ready
			iState:=10;//go go
		ELSIF xEnable AND Axis.StatusWord.1 AND Axis.Modes_of_operation_display <> 8 THEN//need switch mode
			Axis.ControlWord.3:=FALSE;//drop down operation enabled, motor could free move
			iState:=10;
		ELSIF xSimulation THEN
			iState:=20;
		ELSIF xEnable THEN
			iState:=999;//error
		END_IF
	10://Set Mode
		Axis.Modes_of_operation:=8;//Cyclic Synchronous Position Mode
		Axis.ControlWord.3:=Axis.Modes_of_operation_display=8;//Success change mode, enable operation
		otg.CurrentPosition:=DINT_TO_LREAL(Axis.Position_Actual_Value) / lrScale;//Write actual position to otg
		IF Axis.StatusWord.2 AND Axis.Modes_of_operation_display = 8 THEN//Operation Enabled, Mode Changed success
			iState:=20;
		END_IF
	20://Movement
		otg(
			ControlInterface:= FALSE ,
			TargetPosition:= TargetPosition ,
			TargetVelocity:= 0 ,
			CycleTime:= CycleTime,
			MaxVelocity:= MaxVelocity ,
			MaxAcceleration:= MaxAcceleration ,
			MaxJerk:= MaxJerk);//accept new position and going on

		IF otg.NewPosition >= 0 THEN
			Axis.Target_Position := LREAL_TO_DINT(otg.NewPosition * lrScale);
		ELSE
			Axis.Target_Position := - LREAL_TO_DINT( - otg.NewPosition * lrScale);//it fix negative overflow problem.
		END_IF

		IF Axis.StatusWord.13 OR Axis.StatusWord.3 OR otg.xError THEN//Axis Error
			iState:=999;
		ELSIF NOT xEnable THEN
			iState:=0;
		END_IF
	999://Error wait
		xError:=TRUE;
		IF NOT xEnable THEN
			iState:=0;
		END_IF
END_CASE

END_FUNCTION_BLOCK

(* ---- opensml_sync_velocity.st ---- *)
(*
 * OpenSML Cyclic Synchronous Velocity via S7RTT OTG (streams position in mode 8).
 * Vendored from OpenSML (https://github.com/feecat/OpenSML), GPL-3.0.
 *)
FUNCTION_BLOCK OpenSML_SyncVelocity
VAR_IN_OUT
	Axis:OpenSML_Axis;
END_VAR
VAR_INPUT
	MaxVelocity :LREAL:=2000;
	MaxAcceleration :LREAL:=200;
	MaxJerk :LREAL:=200;
	CycleTime:LREAL:=0.001;//0.001 = 1ms

	TargetVelocity :LREAL;
	xEnable: BOOL;
	lrScale:LREAL:=1.0;
	xSimulation: BOOL;
END_VAR
VAR_OUTPUT
	xError: BOOL;
END_VAR
VAR
	otg : FB_S7RTT_OTG;
	iState:INT;

END_VAR

(*
Normally we use CSP(=8) as CSV(=9) cus mostly servo dont have TargetVelocity PDO by default.
If you really want use CSV mode, Please connect OpenSML_SyncVelocity.otg.NewVelocity to TargetVelocity PDO after scale.

Cyclic Synchronous Position Mode (=8)
Set 6060(Op mode) and 60C2(Interpolation time period) at Startup Parameters.

#####################################
NEED StruckigLight Library for Quadratic Velocity Ramp Calculate.

If in movement, Please DO NOT Drop down xEnable.
#####################################
*)
CASE iState OF
	0://start
		xError:=FALSE;
		IF xEnable AND Axis.StatusWord.1 AND Axis.StatusWord.2 AND Axis.Modes_of_operation_display = 8 AND NOT Axis.StatusWord.3 THEN//ready
			iState:=10;//go go
		ELSIF xEnable AND Axis.StatusWord.1 AND Axis.Modes_of_operation_display <> 8 THEN//need switch mode
			Axis.ControlWord.3:=FALSE;//drop down operation enabled, motor could free move
			iState:=10;
		ELSIF xSimulation THEN
			iState:=20;
		ELSIF xEnable THEN
			iState:=999;//error
		END_IF
	10://Set Mode
		Axis.Modes_of_operation:=8;//Cyclic Synchronous Position Mode
		Axis.ControlWord.3:=Axis.Modes_of_operation_display=8;//Success change mode, enable operation
		otg.CurrentPosition:=DINT_TO_LREAL(Axis.Position_Actual_Value) / lrScale;//Write actual position to otg
		IF Axis.StatusWord.2 AND Axis.Modes_of_operation_display = 8 THEN//Operation Enabled, Mode Changed success
			iState:=20;
		END_IF
	20://Movement
		otg(
			ControlInterface:= TRUE ,
			TargetPosition:= 0 ,
			TargetVelocity:= TargetVelocity ,
			CycleTime:=CycleTime,
			MaxVelocity:= MaxVelocity ,
			MaxAcceleration:= MaxAcceleration ,
			MaxJerk:= MaxJerk);//accept new velocity and going on

		IF otg.NewPosition >= 0 THEN
			Axis.Target_Position := LREAL_TO_DINT(otg.NewPosition * lrScale);
		ELSE
			Axis.Target_Position := - LREAL_TO_DINT( - otg.NewPosition * lrScale);//it fix negative overflow problem.
		END_IF

		IF Axis.StatusWord.13 OR Axis.StatusWord.3 OR otg.xError THEN//Axis Error
			iState:=999;
		ELSIF NOT xEnable THEN
			iState:=0;
		END_IF
	999://Error wait
		xError:=TRUE;
		IF NOT xEnable THEN
			iState:=0;
		END_IF
END_CASE

END_FUNCTION_BLOCK

(* ---- s7rtt_blocks.st ---- *)
(*
 * S7RTT online trajectory generator: FB_S7RTT_OTG + FB_S7RTT_Plan.
 * Vendored from S7RTT (https://github.com/feecat/S7RTT), Apache-2.0.
 * Converted from PLCopen XML. Single-axis 7-segment S-curve OTG.
 *)

FUNCTION_BLOCK FB_S7RTT_OTG
VAR_INPUT
	ControlInterface : BOOL := FALSE;
	TargetPosition : LREAL;
	TargetVelocity : LREAL := 0;
	CycleTime : LREAL := 0.001;
	MaxVelocity : LREAL := 10;
	MaxAcceleration : LREAL := 10;
	MaxJerk : LREAL := 10;
	CurrentPosition : LREAL;
END_VAR
VAR_OUTPUT
	NewPosition : LREAL;
	NewVelocity : LREAL;
	NewAcceleration : LREAL;
	xError : BOOL;
END_VAR
VAR
	_ControlInterface : BOOL;
	_TargetPosition : LREAL;
	_TargetVelocity : LREAL;
	_CycleTime : LREAL;
	_MaxVelocity : LREAL;
	_MaxAcceleration : LREAL;
	_MaxJerk : LREAL;
	_CurrentPosition : LREAL;
	xExecute : BOOL;
	fbS7Planner : FB_S7RTT_Plan;
	stS7Limits : ST_MotionLimits;
	stS7Start : ST_MotionState;
	stS7Result : ST_MotionState;
	fS7Timer : LREAL;
END_VAR

// check if input changed
IF (ControlInterface <> _ControlInterface) OR
	(TargetPosition <> _TargetPosition) OR
	(TargetVelocity <> _TargetVelocity) OR
	(CycleTime <> _CycleTime) OR
	(MaxVelocity <> _MaxVelocity) OR
	(MaxAcceleration <> _MaxAcceleration) OR
	(MaxJerk <> _MaxJerk) OR
	(CurrentPosition <> _CurrentPosition) THEN

	IF CurrentPosition <> _CurrentPosition THEN
		stS7Start.fPos := CurrentPosition;
		stS7Result.fPos := CurrentPosition;
		_CurrentPosition := CurrentPosition;
	END_IF
	_ControlInterface := ControlInterface;
	_TargetPosition := TargetPosition;
	_TargetVelocity := TargetVelocity;
	_CycleTime := CycleTime;
	_MaxVelocity := MaxVelocity;
	_MaxAcceleration := MaxAcceleration;
	_MaxJerk := MaxJerk;

	xExecute:=TRUE;
END_IF

// main logic
IF xExecute THEN
    stS7Start.fPos := stS7Result.fPos;
    stS7Start.fVel := stS7Result.fVel;
    stS7Start.fAcc := stS7Result.fAcc;
    stS7Start.fDuration := 0.0;

    stS7Limits.fVelMax := MaxVelocity;
    stS7Limits.fAccMax := MaxAcceleration;
    stS7Limits.fJerkMax := MaxJerk;

    fbS7Planner.ModeVelocity := ControlInterface;
    fbS7Planner.StartState := stS7Start;
    fbS7Planner.TargetPos := TargetPosition;
    fbS7Planner.TargetVel := TargetVelocity;
    fbS7Planner.Limits := stS7Limits;

    fS7Timer := 0.0;
END_IF

fbS7Planner(Execute:=xExecute,Error=>xError);

xExecute := FALSE;

fS7Timer := fS7Timer + CycleTime;

stS7Result := FC_S7RTT_AtTime(
	Trajectory := fbS7Planner.Trajectory,
	SegCount := fbS7Planner.SegmentCount,
	ElapsedTime := fS7Timer
);

NewPosition:=stS7Result.fPos;
NewVelocity:=stS7Result.fVel;
NewAcceleration:=stS7Result.fAcc;
END_FUNCTION_BLOCK

FUNCTION_BLOCK FB_S7RTT_Plan
VAR_INPUT
	Execute : BOOL;
	ModeVelocity : BOOL;
	StartState : ST_MotionState;
	TargetPos : LREAL;
	TargetVel : LREAL;
	Limits : ST_MotionLimits;
END_VAR
VAR_OUTPUT
	Done : BOOL;
	Error : BOOL;
	SegmentCount : INT;
	Trajectory : ARRAY[1..32] OF ST_MotionState;
END_VAR
VAR
	trig_exec : BOOL;
	prev_exec : BOOL;
	c_pos : LREAL;
	c_vel : LREAL;
	c_acc : LREAL;
	i : INT;
	k : INT;
	dist_req : LREAL;
	t_rec : LREAL;
	gap : LREAL;
	d_upper : LREAL;
	d_lower : LREAL;
	t_cruise : LREAL;
	iter : INT;
	sa : LREAL;
	sb : LREAL;
	sc : LREAL;
	fa : LREAL;
	fb : LREAL;
	fc : LREAL;
	sd : LREAL;
	se : LREAL;
	tol1 : LREAL;
	xm : LREAL;
	min1 : LREAL;
	min2 : LREAL;
	fCoefP : LREAL;
	fCoefQ : LREAL;
	fCoefR : LREAL;
	fCoefS : LREAL;
	mflag : BOOL;
	use_optimal : BOOL;
	opt_success : BOOL;
	j_idx : INT;
	j_apply : LREAL;
	search_horizon : LREAL;
	t_est : LREAL;
	sim_p : LREAL;
	sim_v : LREAL;
	sim_a : LREAL;
	limit_a : LREAL;
	dist_to_lim : LREAL;
	t_ramp : LREAL;
	t_hold : LREAL;
	sat_dt : LREAL;
	sat_j : LREAL;
	valid_curr : BOOL;
	best_t_curr : LREAL;
	dur_curr : LREAL;
	winner_found : BOOL;
	winner_dur : LREAL;
	winner_t : LREAL;
	winner_j : LREAL;
	best_v : LREAL;
	v_mid : LREAL;
	a_mid : LREAL;
	v_inertial : LREAL;
	d_inertial : LREAL;
	t_to_zero : LREAL;
	j_restore : LREAL;
	t_shape_buf : ARRAY[1..5] OF LREAL;
	j_shape_buf : ARRAY[1..5] OF LREAL;
	shape_cnt : INT;
	ref_idx : INT;
	max_dt : LREAL;
	dt_fix : LREAL;
	v_cruise_start : LREAL;
	EPS_TIME : LREAL := 1E-10;
	EPS_VAL : LREAL := 1E-10;
	EPS_ACC : LREAL := 1E-10;
	EPS_DIST : LREAL := 1E-10;
	MATH_EPS : LREAL := 1E-10;
	SOLVER_TOL : LREAL := 1E-10;
	SOLVER_EPS : LREAL := 2.22E-16;
	SOLVER_COARSE : LREAL := 0.0001;
	MAX_ITER : INT := 50;
END_VAR

// ==============================================================================
// File Name:    FB_S7RTT_Plan.st
// Author:       feecat
// Version:      V1.8.1
// Description:  Simple 7seg Real-Time Trajectory Generator
// Website:      https://github.com/feecat/S7RTT
// License:      Apache License Version 2.0
// ==============================================================================
//
// Licensed under the Apache License, Version 2.0 (the "License");
// you may not use this file except in compliance with the License.
// You may obtain a copy of the License at
//
//     http://www.apache.org/licenses/LICENSE-2.0
//
// Unless required by applicable law or agreed to in writing, software
// distributed under the License is distributed on an "AS IS" BASIS,
// WITHOUT WARRANTIES OR CONDITIONS OF ANY KIND, either express or implied.
// See the License for the specific language governing permissions and
// limitations under the License.
// ==============================================================================

trig_exec := Execute AND NOT prev_exec;
prev_exec := Execute;

IF NOT Execute THEN
	Done := FALSE; Error := FALSE; RETURN;
END_IF

IF NOT trig_exec THEN RETURN; END_IF;

// --- Initialization ---
Done := FALSE;
Error := FALSE;
SegmentCount := 0;
opt_success := FALSE;

IF Limits.fVelMax <= 0.0 OR Limits.fAccMax <= 0.0 OR Limits.fJerkMax <= 0.0 THEN
	Error := TRUE; RETURN;
END_IF;

c_pos := StartState.fPos; c_vel := StartState.fVel; c_acc := StartState.fAcc;

// ========================================================
// 1. Acceleration Recovery (Safety Decel)
// ========================================================
IF c_acc > Limits.fAccMax + EPS_ACC THEN
	// Positive Saturation: Accel is too high positive, must reduce
	j_restore := -Limits.fJerkMax;
	limit_a := Limits.fAccMax;
	t_rec := (c_acc - limit_a) / (-j_restore);

	IF t_rec > EPS_TIME THEN
		SegmentCount := SegmentCount + 1;
		Trajectory[SegmentCount].fDuration := t_rec;
		Trajectory[SegmentCount].fJerk     := j_restore;
		// Integ State
		c_pos := c_pos + c_vel * t_rec + 0.5 * c_acc * t_rec*t_rec + (1.0/6.0) * j_restore * t_rec*t_rec*t_rec;
		c_vel := c_vel + c_acc * t_rec + 0.5 * j_restore * t_rec*t_rec;
		c_acc := limit_a;
	END_IF;

ELSIF c_acc < -Limits.fAccMax - EPS_ACC THEN
	// Negative Saturation: Accel is too low negative, must increase
	j_restore := Limits.fJerkMax;
	limit_a := -Limits.fAccMax;
	t_rec := (c_acc - limit_a) / (-j_restore); // Note: -j_restore here implies dividing by -JerkMax which is negative

	IF t_rec > EPS_TIME THEN
		SegmentCount := SegmentCount + 1;
		Trajectory[SegmentCount].fDuration := t_rec;
		Trajectory[SegmentCount].fJerk     := j_restore;
		// Integ State
		c_pos := c_pos + c_vel * t_rec + 0.5 * c_acc * t_rec*t_rec + (1.0/6.0) * j_restore * t_rec*t_rec*t_rec;
		c_vel := c_vel + c_acc * t_rec + 0.5 * j_restore * t_rec*t_rec;
		c_acc := limit_a;
	END_IF;
END_IF;

// ========================================================
// 2. Plan Generation
// ========================================================
IF ModeVelocity THEN
	// --- Velocity Mode (Unchanged Logic, New Constants) ---
	v_mid := TargetVel;
	IF v_mid > Limits.fVelMax THEN v_mid := Limits.fVelMax; END_IF;
	IF v_mid < -Limits.fVelMax THEN v_mid := -Limits.fVelMax; END_IF;

	shape_cnt := FC_S7RTT_BuildProfile(c_vel, c_acc, v_mid, Limits.fAccMax, Limits.fJerkMax, t_shape_buf, j_shape_buf);
	IF shape_cnt > 0 THEN
		FOR i := 1 TO shape_cnt DO
			IF SegmentCount < 32 THEN
				SegmentCount := SegmentCount + 1;
				Trajectory[SegmentCount].fDuration := t_shape_buf[i];
				Trajectory[SegmentCount].fJerk     := j_shape_buf[i];
			END_IF;
		END_FOR;
	ELSE
		FOR i := 1 TO 31 DO
			SegmentCount := SegmentCount + 1;
			Trajectory[SegmentCount].fDuration := 0;
			Trajectory[SegmentCount].fJerk     := 0;
		END_FOR;
	END_IF
ELSE
	// --- Position Mode ---
	dist_req := TargetPos - c_pos;

	// Capacity Check (Can we reach target without hitting velocity limits?)
	// Note: FC_S7RTT_CalcTrajDist returns distance traveled to reach TargetVel via +/- VelMax
	d_upper := FC_S7RTT_CalcTrajDist(Limits.fVelMax, c_vel, c_acc, TargetVel, Limits.fAccMax, Limits.fJerkMax);
	d_lower := FC_S7RTT_CalcTrajDist(-Limits.fVelMax, c_vel, c_acc, TargetVel, Limits.fAccMax, Limits.fJerkMax);

	// Decision: Cruise or Optimal?
	use_optimal := TRUE;
	IF dist_req > d_upper + EPS_DIST THEN use_optimal := FALSE; END_IF;
	IF dist_req < d_lower - EPS_DIST THEN use_optimal := FALSE; END_IF;

	// ========================================================
	// 2.1 Time Optimal Solver (New V1.7 Feature)
	// ========================================================
	IF use_optimal THEN
		winner_found := FALSE;
		winner_dur := 1.0E10; // Init Large

		// Estimate search horizon
		t_est := (ABS(c_vel) + Limits.fVelMax) / Limits.fAccMax;
		IF t_est < 1.0 THEN t_est := 1.0; END_IF;
		search_horizon := t_est * 2.0 + 5.0;

		// Bidirectional Competition: Try +Jerk and -Jerk
		FOR j_idx := 0 TO 1 DO
			IF j_idx = 0 THEN j_apply := Limits.fJerkMax; ELSE j_apply := -Limits.fJerkMax; END_IF;
			valid_curr := FALSE;

			// Brent Solver Setup: Range [0, search_horizon]
			sa := 0.0; sb := search_horizon;

			// --- Evaluate at sa (0.0) ---
			// Inline Simulation Block 1
			sim_p := c_pos; sim_v := c_vel; sim_a := c_acc; // Reset State
			// Integrate Saturated (t=0 -> no effect), then Build Profile
			shape_cnt := FC_S7RTT_BuildProfile(sim_v, sim_a, TargetVel, Limits.fAccMax, Limits.fJerkMax, t_shape_buf, j_shape_buf);
			FOR k:=1 TO shape_cnt DO
				sim_p := sim_p + sim_v*t_shape_buf[k] + 0.5*sim_a*t_shape_buf[k]*t_shape_buf[k] + (1.0/6.0)*j_shape_buf[k]*t_shape_buf[k]*t_shape_buf[k]*t_shape_buf[k];
				sim_v := sim_v + sim_a*t_shape_buf[k] + 0.5*j_shape_buf[k]*t_shape_buf[k]*t_shape_buf[k];
				sim_a := sim_a + j_shape_buf[k]*t_shape_buf[k];
			END_FOR;
			fa := sim_p - TargetPos; // Error at t=0

			IF ABS(fa) < SOLVER_COARSE THEN
				best_t_curr := 0.0; valid_curr := TRUE;
			ELSE
				// --- Evaluate at sb (horizon) ---
				// Inline Simulation Block 2
				sim_p := c_pos; sim_v := c_vel; sim_a := c_acc;
				limit_a := Limits.fAccMax; IF j_apply < 0 THEN limit_a := -Limits.fAccMax; END_IF;
				dist_to_lim := limit_a - sim_a;
				IF (j_apply > 0 AND dist_to_lim > -MATH_EPS) OR (j_apply < 0 AND dist_to_lim < MATH_EPS) THEN t_ramp := dist_to_lim / j_apply; ELSE t_ramp := 0.0; END_IF;
				// Saturated Int (simplified logic for end of range)
				IF sb <= t_ramp THEN
					sim_p:=sim_p+sim_v*sb+0.5*sim_a*sb*sb+(1.0/6.0)*j_apply*sb*sb*sb; sim_v:=sim_v+sim_a*sb+0.5*j_apply*sb*sb; sim_a:=sim_a+j_apply*sb;
				ELSE
					sim_p:=sim_p+sim_v*t_ramp+0.5*sim_a*t_ramp*t_ramp+(1.0/6.0)*j_apply*t_ramp*t_ramp*t_ramp; sim_v:=sim_v+sim_a*t_ramp+0.5*j_apply*t_ramp*t_ramp; sim_a:=sim_a+j_apply*t_ramp;
					sim_a:=limit_a; t_hold:=sb-t_ramp;
					sim_p:=sim_p+sim_v*t_hold+0.5*sim_a*t_hold*t_hold; sim_v:=sim_v+sim_a*t_hold;
				END_IF;
				shape_cnt := FC_S7RTT_BuildProfile(sim_v, sim_a, TargetVel, Limits.fAccMax, Limits.fJerkMax, t_shape_buf, j_shape_buf);
				FOR k:=1 TO shape_cnt DO sim_p:=sim_p+sim_v*t_shape_buf[k]+0.5*sim_a*t_shape_buf[k]*t_shape_buf[k]+(1.0/6.0)*j_shape_buf[k]*t_shape_buf[k]*t_shape_buf[k]*t_shape_buf[k]; sim_v:=sim_v+sim_a*t_shape_buf[k]+0.5*j_shape_buf[k]*t_shape_buf[k]*t_shape_buf[k]; sim_a:=sim_a+j_shape_buf[k]*t_shape_buf[k]; END_FOR;
				fb := sim_p - TargetPos;

				// Bounds Check
				IF fa * fb <= 0.0 THEN
					// Brent Loop
					sc := sa; fc := fa; sd := sb - sa; se := sd; mflag := TRUE;
					FOR iter := 1 TO MAX_ITER DO
						IF ABS(fc) < ABS(fb) THEN sa:=sb; sb:=sc; sc:=sa; fa:=fb; fb:=fc; fc:=fa; END_IF;
						tol1 := 2.0 * SOLVER_EPS * ABS(sb) + 0.5 * SOLVER_TOL; xm := 0.5 * (sc - sb);
						IF ABS(xm) <= tol1 OR fb = 0.0 THEN EXIT; END_IF;
						IF ABS(se) >= tol1 AND ABS(fa) > ABS(fb) THEN
							fCoefS := fb / fa;
							IF sa = sc THEN fCoefP := 2.0*xm*fCoefS; fCoefQ := 1.0-fCoefS;
							ELSE fCoefQ := fa/fc; fCoefR := fb/fc; fCoefP := fCoefS*(2.0*xm*fCoefQ*(fCoefQ-fCoefR)-(sb-sa)*(fCoefR-1.0)); fCoefQ := (fCoefQ-1.0)*(fCoefR-1.0)*(fCoefS-1.0); END_IF;
							IF fCoefP > 0.0 THEN fCoefQ := -fCoefQ; END_IF; fCoefP := ABS(fCoefP);
							min1 := 3.0*xm*fCoefQ - ABS(tol1*fCoefQ); min2 := ABS(se*fCoefQ);
							IF 2.0*fCoefP < min1 THEN
								IF mflag THEN IF 2.0*fCoefP < min2 THEN se:=sd; sd:=fCoefP/fCoefQ; mflag:=FALSE; ELSE sd:=xm; se:=sd; mflag:=TRUE; END_IF;
								ELSE IF 2.0*fCoefP < ABS(sd*fCoefQ) THEN se:=sd; sd:=fCoefP/fCoefQ; mflag:=FALSE; ELSE sd:=xm; se:=sd; mflag:=TRUE; END_IF; END_IF;
							ELSE sd:=xm; se:=sd; mflag:=TRUE; END_IF;
						ELSE sd:=xm; se:=sd; mflag:=TRUE; END_IF;
						sa := sb; fa := fb;
						IF ABS(sd) > tol1 THEN sb:=sb+sd; ELSE IF xm > 0.0 THEN sb:=sb+tol1; ELSE sb:=sb-tol1; END_IF; END_IF;

						// --- Eval Function (t = sb) ---
						// Only necessary to update fb. Re-use simulation logic.
						sim_p := c_pos; sim_v := c_vel; sim_a := c_acc;
						limit_a := Limits.fAccMax; IF j_apply < 0 THEN limit_a := -Limits.fAccMax; END_IF;
						dist_to_lim := limit_a - sim_a;
						IF (j_apply > 0 AND dist_to_lim > -MATH_EPS) OR (j_apply < 0 AND dist_to_lim < MATH_EPS) THEN t_ramp := dist_to_lim / j_apply; ELSE t_ramp := 0.0; END_IF;
						IF sb <= t_ramp THEN
							IF sb > EPS_TIME THEN sim_p:=sim_p+sim_v*sb+0.5*sim_a*sb*sb+(1.0/6.0)*j_apply*sb*sb*sb; sim_v:=sim_v+sim_a*sb+0.5*j_apply*sb*sb; sim_a:=sim_a+j_apply*sb; END_IF;
						ELSE
							IF t_ramp > EPS_TIME THEN sim_p:=sim_p+sim_v*t_ramp+0.5*sim_a*t_ramp*t_ramp+(1.0/6.0)*j_apply*t_ramp*t_ramp*t_ramp; sim_v:=sim_v+sim_a*t_ramp+0.5*j_apply*t_ramp*t_ramp; sim_a:=sim_a+j_apply*t_ramp; END_IF;
							sim_a:=limit_a; t_hold:=sb-t_ramp;
							IF t_hold > EPS_TIME THEN sim_p:=sim_p+sim_v*t_hold+0.5*sim_a*t_hold*t_hold; sim_v:=sim_v+sim_a*t_hold; END_IF;
						END_IF;
						shape_cnt := FC_S7RTT_BuildProfile(sim_v, sim_a, TargetVel, Limits.fAccMax, Limits.fJerkMax, t_shape_buf, j_shape_buf);
						FOR k:=1 TO shape_cnt DO sim_p:=sim_p+sim_v*t_shape_buf[k]+0.5*sim_a*t_shape_buf[k]*t_shape_buf[k]+(1.0/6.0)*j_shape_buf[k]*t_shape_buf[k]*t_shape_buf[k]*t_shape_buf[k]; sim_v:=sim_v+sim_a*t_shape_buf[k]+0.5*j_shape_buf[k]*t_shape_buf[k]*t_shape_buf[k]; sim_a:=sim_a+j_shape_buf[k]*t_shape_buf[k]; END_FOR;
						fb := sim_p - TargetPos;
						// --- End Eval ---

						IF (fb > 0.0 AND fc > 0.0) OR (fb < 0.0 AND fc < 0.0) THEN sc := sa; fc := fa; sd := sb - sa; se := sd; mflag := TRUE; END_IF;
					END_FOR;
					best_t_curr := sb;
					IF ABS(fb) <= SOLVER_COARSE THEN valid_curr := TRUE; END_IF;
				END_IF;
			END_IF;

			// Calculate Total Duration for Comparison
			IF valid_curr THEN
				dur_curr := 0.0;
				// Saturated Time
				limit_a := Limits.fAccMax; IF j_apply < 0 THEN limit_a := -Limits.fAccMax; END_IF;
				dist_to_lim := limit_a - c_acc;
				IF (j_apply > 0 AND dist_to_lim > -MATH_EPS) OR (j_apply < 0 AND dist_to_lim < MATH_EPS) THEN t_ramp := dist_to_lim / j_apply; ELSE t_ramp := 0.0; END_IF;
				IF best_t_curr <= t_ramp THEN dur_curr := best_t_curr;
				ELSE dur_curr := best_t_curr; // t_ramp + (t - t_ramp)
				END_IF;
				// Sim to get intermediate state for remaining profile
				sim_p := c_pos; sim_v := c_vel; sim_a := c_acc;
				IF best_t_curr <= t_ramp THEN
					IF best_t_curr > EPS_TIME THEN sim_v:=sim_v+sim_a*best_t_curr+0.5*j_apply*best_t_curr*best_t_curr; sim_a:=sim_a+j_apply*best_t_curr; END_IF;
				ELSE
					IF t_ramp > EPS_TIME THEN sim_v:=sim_v+sim_a*t_ramp+0.5*j_apply*t_ramp*t_ramp; sim_a:=sim_a+j_apply*t_ramp; END_IF;
					sim_a:=limit_a; t_hold:=best_t_curr-t_ramp;
					IF t_hold > EPS_TIME THEN sim_v:=sim_v+sim_a*t_hold; END_IF;
				END_IF;
				shape_cnt := FC_S7RTT_BuildProfile(sim_v, sim_a, TargetVel, Limits.fAccMax, Limits.fJerkMax, t_shape_buf, j_shape_buf);
				FOR k:=1 TO shape_cnt DO dur_curr := dur_curr + t_shape_buf[k]; END_FOR;

				// Update Winner
				IF dur_curr < winner_dur THEN winner_dur := dur_curr; winner_t := best_t_curr; winner_j := j_apply; winner_found := TRUE; END_IF;
			END_IF;
		END_FOR;

		// Construct Winner
		IF winner_found THEN
			opt_success := TRUE;
			limit_a := Limits.fAccMax; IF winner_j < 0 THEN limit_a := -Limits.fAccMax; END_IF;
			dist_to_lim := limit_a - c_acc;
			IF (winner_j > 0 AND dist_to_lim > -MATH_EPS) OR (winner_j < 0 AND dist_to_lim < MATH_EPS) THEN t_ramp := dist_to_lim / winner_j; ELSE t_ramp := 0.0; END_IF;

			IF winner_t <= t_ramp THEN
				IF winner_t > EPS_TIME THEN
					IF SegmentCount < 32 THEN SegmentCount:=SegmentCount+1; Trajectory[SegmentCount].fDuration:=winner_t; Trajectory[SegmentCount].fJerk:=winner_j; END_IF;
					c_pos:=c_pos+c_vel*winner_t+0.5*c_acc*winner_t*winner_t+(1.0/6.0)*winner_j*winner_t*winner_t*winner_t; c_vel:=c_vel+c_acc*winner_t+0.5*winner_j*winner_t*winner_t; c_acc:=c_acc+winner_j*winner_t;
				END_IF;
			ELSE
				IF t_ramp > EPS_TIME THEN
					IF SegmentCount < 32 THEN SegmentCount:=SegmentCount+1; Trajectory[SegmentCount].fDuration:=t_ramp; Trajectory[SegmentCount].fJerk:=winner_j; END_IF;
					c_pos:=c_pos+c_vel*t_ramp+0.5*c_acc*t_ramp*t_ramp+(1.0/6.0)*winner_j*t_ramp*t_ramp*t_ramp; c_vel:=c_vel+c_acc*t_ramp+0.5*winner_j*t_ramp*t_ramp; c_acc:=c_acc+winner_j*t_ramp;
				END_IF;
				c_acc := limit_a; t_hold := winner_t - t_ramp;
				IF t_hold > EPS_TIME THEN
					IF SegmentCount < 32 THEN SegmentCount:=SegmentCount+1; Trajectory[SegmentCount].fDuration:=t_hold; Trajectory[SegmentCount].fJerk:=0.0; END_IF;
					c_pos:=c_pos+c_vel*t_hold+0.5*c_acc*t_hold*t_hold; c_vel:=c_vel+c_acc*t_hold;
				END_IF;
			END_IF;
			shape_cnt := FC_S7RTT_BuildProfile(c_vel, c_acc, TargetVel, Limits.fAccMax, Limits.fJerkMax, t_shape_buf, j_shape_buf);
			FOR i:=1 TO shape_cnt DO IF SegmentCount < 32 THEN SegmentCount:=SegmentCount+1; Trajectory[SegmentCount].fDuration:=t_shape_buf[i]; Trajectory[SegmentCount].fJerk:=j_shape_buf[i]; END_IF; END_FOR;
		END_IF;
	END_IF;

	// ========================================================
	// 2.2 Fallback / Cruise Logic (Original + Cruise)
	// ========================================================
	IF NOT opt_success THEN
		// If dist_req > d_upper, we Cruise at VMax. If < d_lower, at -VMax.
		// Otherwise, we solve for intermediate peak.

		IF dist_req > d_upper + EPS_DIST THEN best_v := Limits.fVelMax;
		ELSIF dist_req < d_lower - EPS_DIST THEN best_v := -Limits.fVelMax;
		ELSE
			// Bisection Solver (Original Logic, compacted)
			sa := -Limits.fVelMax; sb := Limits.fVelMax;
			// Calc Fa/Fb using helper function logic (Dist via profile)
			// Note: Assuming FC_S7RTT_CalcTrajDist calculates distance for a profile peaking at 'sa'/'sb' then going to TargetVel
			fa := FC_S7RTT_CalcTrajDist(sa, c_vel, c_acc, TargetVel, Limits.fAccMax, Limits.fJerkMax) - dist_req;
			fb := FC_S7RTT_CalcTrajDist(sb, c_vel, c_acc, TargetVel, Limits.fAccMax, Limits.fJerkMax) - dist_req;

			IF fa * fb > 0.0 THEN IF ABS(fa) < ABS(fb) THEN best_v := sa; ELSE best_v := sb; END_IF;
			ELSE
				sc:=sa; fc:=fa; sd:=sb-sa; se:=sd; mflag:=TRUE;
				FOR iter := 1 TO MAX_ITER DO
					IF ABS(fc) < ABS(fb) THEN sa:=sb; sb:=sc; sc:=sa; fa:=fb; fb:=fc; fc:=fa; END_IF;
					tol1 := 2.0 * SOLVER_EPS * ABS(sb) + 0.5 * SOLVER_TOL; xm := 0.5 * (sc - sb);
					IF ABS(xm) <= tol1 OR fb = 0.0 THEN EXIT; END_IF;
					IF ABS(se) >= tol1 AND ABS(fa) > ABS(fb) THEN
						fCoefS := fb/fa;
						IF sa=sc THEN fCoefP:=2.0*xm*fCoefS; fCoefQ:=1.0-fCoefS; ELSE fCoefQ:=fa/fc; fCoefR:=fb/fc; fCoefP:=fCoefS*(2.0*xm*fCoefQ*(fCoefQ-fCoefR)-(sb-sa)*(fCoefR-1.0)); fCoefQ:=(fCoefQ-1.0)*(fCoefR-1.0)*(fCoefS-1.0); END_IF;
						IF fCoefP > 0.0 THEN fCoefQ:=-fCoefQ; END_IF; fCoefP:=ABS(fCoefP); min1:=3.0*xm*fCoefQ-ABS(tol1*fCoefQ); min2:=ABS(se*fCoefQ);
						IF 2.0*fCoefP < min1 THEN IF mflag THEN IF 2.0*fCoefP < min2 THEN se:=sd; sd:=fCoefP/fCoefQ; mflag:=FALSE; ELSE sd:=xm; se:=sd; mflag:=TRUE; END_IF; ELSE IF 2.0*fCoefP < ABS(sd*fCoefQ) THEN se:=sd; sd:=fCoefP/fCoefQ; mflag:=FALSE; ELSE sd:=xm; se:=sd; mflag:=TRUE; END_IF; END_IF; ELSE sd:=xm; se:=sd; mflag:=TRUE; END_IF;
					ELSE sd:=xm; se:=sd; mflag:=TRUE; END_IF;
					sa:=sb; fa:=fb; IF ABS(sd) > tol1 THEN sb:=sb+sd; ELSE IF xm > 0.0 THEN sb:=sb+tol1; ELSE sb:=sb-tol1; END_IF; END_IF;
					fb := FC_S7RTT_CalcTrajDist(sb, c_vel, c_acc, TargetVel, Limits.fAccMax, Limits.fJerkMax) - dist_req;
					IF (fb > 0.0 AND fc > 0.0) OR (fb < 0.0 AND fc < 0.0) THEN sc:=sa; fc:=fa; sd:=sb-sa; se:=sd; mflag:=TRUE; END_IF;
				END_FOR;
				best_v := sb;
			END_IF;
		END_IF;

		// Generate fallback profile
		shape_cnt := FC_S7RTT_BuildProfile(c_vel, c_acc, best_v, Limits.fAccMax, Limits.fJerkMax, t_shape_buf, j_shape_buf);
		FOR i:=1 TO shape_cnt DO
			IF SegmentCount < 32 THEN SegmentCount:=SegmentCount+1; Trajectory[SegmentCount].fDuration:=t_shape_buf[i]; Trajectory[SegmentCount].fJerk:=j_shape_buf[i]; END_IF;
			c_pos:=c_pos+c_vel*t_shape_buf[i]+0.5*c_acc*t_shape_buf[i]*t_shape_buf[i]+(1.0/6.0)*j_shape_buf[i]*t_shape_buf[i]*t_shape_buf[i]*t_shape_buf[i];
			c_vel:=c_vel+c_acc*t_shape_buf[i]+0.5*j_shape_buf[i]*t_shape_buf[i]*t_shape_buf[i]; c_acc:=c_acc+j_shape_buf[i]*t_shape_buf[i];
		END_FOR;
		// Add Cruise if needed (gap logic)
		c_acc := 0.0;
		// Sim fwd
		sim_p := c_pos; sim_v := c_vel; sim_a := 0.0;
		shape_cnt := FC_S7RTT_BuildProfile(sim_v, sim_a, TargetVel, Limits.fAccMax, Limits.fJerkMax, t_shape_buf, j_shape_buf);
		FOR k:=1 TO shape_cnt DO sim_p:=sim_p+sim_v*t_shape_buf[k]+0.5*sim_a*t_shape_buf[k]*t_shape_buf[k]+(1.0/6.0)*j_shape_buf[k]*t_shape_buf[k]*t_shape_buf[k]*t_shape_buf[k]; sim_v:=sim_v+sim_a*t_shape_buf[k]+0.5*j_shape_buf[k]*t_shape_buf[k]*t_shape_buf[k]; sim_a:=sim_a+j_shape_buf[k]*t_shape_buf[k]; END_FOR;
		gap := TargetPos - sim_p;
		IF ABS(c_vel) > EPS_VAL AND ABS(gap) > EPS_DIST THEN
			t_cruise := gap / c_vel;
			IF t_cruise > EPS_TIME THEN
				IF SegmentCount < 32 THEN SegmentCount:=SegmentCount+1; Trajectory[SegmentCount].fDuration:=t_cruise; Trajectory[SegmentCount].fJerk:=0.0; END_IF;
				c_pos := c_pos + c_vel * t_cruise;
			END_IF;
		END_IF;
		// Final Decel
		shape_cnt := FC_S7RTT_BuildProfile(c_vel, c_acc, TargetVel, Limits.fAccMax, Limits.fJerkMax, t_shape_buf, j_shape_buf);
		FOR i:=1 TO shape_cnt DO IF SegmentCount < 32 THEN SegmentCount:=SegmentCount+1; Trajectory[SegmentCount].fDuration:=t_shape_buf[i]; Trajectory[SegmentCount].fJerk:=j_shape_buf[i]; END_IF; END_FOR;
	END_IF;
END_IF;

// ========================================================
// 2.5 Trajectory Refinement (Precision Fix)
// ========================================================
IF SegmentCount > 0 AND NOT ModeVelocity THEN
	c_pos := StartState.fPos; c_vel := StartState.fVel; c_acc := StartState.fAcc;
	ref_idx := -1; max_dt := -1.0;
	FOR i := 1 TO SegmentCount DO
		t_rec := Trajectory[i].fDuration; j_restore := Trajectory[i].fJerk;
		IF ABS(j_restore) < MATH_EPS AND ABS(c_acc) < EPS_ACC THEN IF t_rec > max_dt THEN max_dt:=t_rec; ref_idx:=i; v_cruise_start:=c_vel; END_IF; END_IF;
		c_pos:=c_pos+c_vel*t_rec+0.5*c_acc*t_rec*t_rec+(1.0/6.0)*j_restore*t_rec*t_rec*t_rec; c_vel:=c_vel+c_acc*t_rec+0.5*j_restore*t_rec*t_rec; c_acc:=c_acc+j_restore*t_rec;
	END_FOR;
	gap := TargetPos - c_pos;
	IF ref_idx <> -1 AND ABS(gap) > EPS_DIST AND ABS(v_cruise_start) > EPS_VAL THEN
		dt_fix := gap / v_cruise_start;
		Trajectory[ref_idx].fDuration := Trajectory[ref_idx].fDuration + dt_fix;
		IF Trajectory[ref_idx].fDuration < EPS_TIME THEN Trajectory[ref_idx].fDuration := EPS_TIME; END_IF;
	END_IF;
END_IF;

// ========================================================
// 3. Final Pass
// ========================================================
c_pos := StartState.fPos; c_vel := StartState.fVel; c_acc := StartState.fAcc;
FOR i := 1 TO SegmentCount DO
	Trajectory[i].fPos := c_pos; Trajectory[i].fVel := c_vel; Trajectory[i].fAcc := c_acc;
	t_rec := Trajectory[i].fDuration; j_restore := Trajectory[i].fJerk;
	c_pos:=c_pos+c_vel*t_rec+0.5*c_acc*t_rec*t_rec+(1.0/6.0)*j_restore*t_rec*t_rec*t_rec; c_vel:=c_vel+c_acc*t_rec+0.5*j_restore*t_rec*t_rec; c_acc:=c_acc+j_restore*t_rec;
END_FOR;

IF SegmentCount = 0 THEN
	Trajectory[1]:= StartState;
	Trajectory[1].fDuration := 0; Trajectory[1].fJerk := 0; Trajectory[1].fAcc := 0;
	SegmentCount := 1;
END_IF

Done := TRUE;
Done := TRUE;
END_FUNCTION_BLOCK

(* ---- sm3_drive.st ---- *)
(*
 * SM_Drive_GenericDS402 — generic CiA 402 (DS402) drive bridge.
 *
 * The OpenPLC analogue of CODESYS SM_Drive_ETC_GenericDSP402. One instance per
 * axis, called once per scan (generated by the editor at the top of the scan).
 * It is the ONLY block that copies the CiA 402 PDO image and converts between
 * increments and technical units. Data flow forms a one-scan pipeline:
 *   - copy this scan's drive TxPDO inputs  -> Axis.Drive + engineering feedback
 *   - copy last scan's MC_* command words  -> drive RxPDO outputs
 * The MC_* blocks run in between and act on Axis / Axis.Drive.
 *)
FUNCTION_BLOCK SM_Drive_GenericDS402
VAR_IN_OUT
	Axis : AXIS_REF_SM3;
END_VAR
VAR_INPUT
	(* from drive TxPDOs *)
	wStatusWord : UINT;                    (* 0x6041 *)
	siModesDisplay : SINT;                 (* 0x6061 *)
	diActualPosition : DINT;               (* 0x6064 *)
	diActualVelocity : DINT;               (* 0x606C *)
	iActualTorque : INT;                   (* 0x6077 *)
	bOnline : BOOL := TRUE;                (* fieldbus/slave operational *)
END_VAR
VAR_OUTPUT
	(* to drive RxPDOs *)
	wControlWord : UINT;                   (* 0x6040 *)
	siModes : SINT;                        (* 0x6060 *)
	diTargetPosition : DINT;               (* 0x607A *)
	udiProfileVelocity : UDINT;            (* 0x6081 *)
	diTargetVelocity : DINT;               (* 0x60FF *)
	iTargetTorque : INT;                   (* 0x6071 *)
END_VAR

(* ---- 1. Ingest drive feedback into the raw CiA 402 image ---- *)
Axis.Drive.StatusWord := wStatusWord;
Axis.Drive.Modes_of_operation_display := siModesDisplay;
Axis.Drive.Position_Actual_Value := diActualPosition;
Axis.Drive.Velocity_Actual_Value := diActualVelocity;
Axis.Drive.Torque_Actual_Value := iActualTorque;

(* ---- 2. Refresh the increments<->units scale factor ---- *)
IF Axis.dwRatioTechUnitsDenom = DWORD#0 THEN
	Axis.dwRatioTechUnitsDenom := DWORD#1;
END_IF
Axis.fIncPerUnit := Axis.fScalefactor
	* DINT_TO_LREAL(Axis.iRatioTechUnitsNum)
	/ DWORD_TO_LREAL(Axis.dwRatioTechUnitsDenom);
IF Axis.fIncPerUnit = 0.0 THEN
	Axis.fIncPerUnit := 1.0;
END_IF

(* ---- 3. Engineering-unit feedback ---- *)
Axis.fActPosition := DINT_TO_LREAL(Axis.Drive.Position_Actual_Value) / Axis.fIncPerUnit;
Axis.fActVelocity := DINT_TO_LREAL(Axis.Drive.Velocity_Actual_Value) / Axis.fIncPerUnit;
Axis.fActTorque := INT_TO_LREAL(Axis.Drive.Torque_Actual_Value);
Axis.byRealControllerMode := SINT_TO_BYTE(Axis.Drive.Modes_of_operation_display);

(* ---- 4. Communication + error + PLCopen state ---- *)
Axis.bCommunication := bOnline;
Axis.wCommunicationState := UINT_TO_WORD(Axis.Drive.StatusWord);
Axis.bRegulatorRealState := Axis.Drive.StatusWord.2;   (* Operation enabled *)
Axis.bDriveStartRealState := NOT Axis.Drive.StatusWord.5; (* NOT quick-stop-active *)
Axis.bError := Axis.Drive.StatusWord.3;                (* Fault *)

IF NOT bOnline THEN
	Axis.dwErrorID := DWORD#1;      (* SMC_DI_GENERAL_COMMUNICATION_ERROR *)
	Axis.nAxisState := SMC_AXIS_STATE.errorstop;
ELSIF Axis.bError THEN
	Axis.dwErrorID := DWORD#2;      (* SMC_DI_AXIS_ERROR *)
	Axis.nAxisState := SMC_AXIS_STATE.errorstop;
ELSE
	Axis.dwErrorID := DWORD#0;      (* SMC_NO_ERROR *)
	IF NOT Axis.Drive.StatusWord.2 THEN
		Axis.nAxisState := SMC_AXIS_STATE.power_off;        (* not operation-enabled *)
	ELSIF Axis.Drive.StatusWord.14 THEN
		Axis.nAxisState := SMC_AXIS_STATE.standstill;       (* SW bit14: standstill *)
	ELSIF Axis.Drive.Modes_of_operation_display = 3 THEN
		Axis.nAxisState := SMC_AXIS_STATE.continuous_motion;(* profile velocity *)
	ELSIF Axis.Drive.Modes_of_operation_display = 6 THEN
		Axis.nAxisState := SMC_AXIS_STATE.homing;
	ELSE
		Axis.nAxisState := SMC_AXIS_STATE.discrete_motion;
	END_IF
END_IF

(* ---- 5. Emit the RxPDO command image ---- *)
wControlWord := Axis.Drive.ControlWord;
siModes := Axis.Drive.Modes_of_operation;
diTargetPosition := Axis.Drive.Target_Position;
udiProfileVelocity := Axis.Drive.Profile_Velocity;
diTargetVelocity := Axis.Drive.Target_Velocity;
iTargetTorque := Axis.Drive.Target_torque;
END_FUNCTION_BLOCK

(* ---- sm3_mc_blocks.st ---- *)
(*
 * PLCopen MC_* function blocks — CODESYS SoftMotion SM3 compatible.
 *
 * Signatures/units match CODESYS SM3_Basic so CODESYS application code ports
 * unmodified: axis is AXIS_REF_SM3 (VAR_IN_OUT), positions/velocities are LREAL
 * technical units, and the standard PLCopen output set is provided. Each block
 * drives the validated OpenSML CiA 402 engine on the axis's embedded raw drive
 * image (Axis.Drive), converting technical units to increments via
 * Axis.fIncPerUnit (maintained by SM_Drive_GenericDS402).
 *
 * Supported buffering model: single active move (BufferMode Aborting). The
 * BufferMode / Direction inputs are accepted for signature compatibility;
 * blending/queuing across multiple concurrently-executing blocks is not
 * modelled. Acceleration/Deceleration/Jerk are recorded on the axis and, in
 * the drive-side profile modes, honoured by the drive's own ramp objects.
 *)

(* ------------------------------------------------------------------ MC_Power *)
FUNCTION_BLOCK MC_Power
VAR_IN_OUT
	Axis : AXIS_REF_SM3;
END_VAR
VAR_INPUT
	Enable : BOOL;
	bRegulatorOn : BOOL := TRUE;   (* enable power stage / closed loop *)
	bDriveStart : BOOL := TRUE;    (* release quick stop *)
END_VAR
VAR_OUTPUT
	Status : BOOL;                 (* axis ready to move (operation enabled) *)
	bRegulatorRealState : BOOL;
	bDriveStartRealState : BOOL;
	Busy : BOOL;
	Error : BOOL;
	ErrorID : SMC_ERROR;
END_VAR
VAR
	_pwr : OpenSML_Power;
END_VAR
	Axis.bRegulatorOn := Enable AND bRegulatorOn;
	Axis.bDriveStart := Enable AND bDriveStart;
	_pwr(Axis := Axis.Drive,
	     xEnable := Enable AND bRegulatorOn,
	     xEmergencyStop := bDriveStart);
	Status := _pwr.xDone;
	bRegulatorRealState := Axis.bRegulatorRealState;
	bDriveStartRealState := Axis.bDriveStartRealState;
	Busy := (Enable AND bRegulatorOn) AND NOT _pwr.xDone AND NOT _pwr.xError;
	Error := _pwr.xError;
	IF _pwr.xError THEN ErrorID := SMC_REGULATOR_OR_START_NOT_SET;
	ELSE ErrorID := SMC_NO_ERROR; END_IF
END_FUNCTION_BLOCK

(* ---------------------------------------------------------- MC_MoveAbsolute *)
FUNCTION_BLOCK MC_MoveAbsolute
VAR_IN_OUT
	Axis : AXIS_REF_SM3;
END_VAR
VAR_INPUT
	Execute : BOOL;
	Position : LREAL;              (* [u] *)
	Velocity : LREAL;             (* [u/s] *)
	Acceleration : LREAL;
	Deceleration : LREAL;
	Jerk : LREAL;
	Direction : MC_DIRECTION := mcd_positive;
	BufferMode : MC_BUFFER_MODE := mcbm_aborting;
END_VAR
VAR_OUTPUT
	Done : BOOL;
	Busy : BOOL;
	Active : BOOL;
	CommandAborted : BOOL;
	Error : BOOL;
	ErrorID : SMC_ERROR;
END_VAR
VAR
	_pp : OpenSML_ProfilePosition;
END_VAR
	IF Execute THEN
		Axis.byControllerMode := BYTE#3;   (* SMC_position *)
		Axis.fSetPosition := Position;
		Axis.fSetVelocity := Velocity;
		Axis.fSetAcceleration := Acceleration;
		Axis.fSetDeceleration := Deceleration;
		Axis.fSetJerk := Jerk;
	END_IF
	_pp(Axis := Axis.Drive,
	    xEnable := Execute,
	    xExecute := Execute,
	    xContinueMove := (BufferMode <> mcbm_aborting),
	    xRelativeMode := FALSE,
	    diTargetPosition := LREAL_TO_DINT(Position * Axis.fIncPerUnit),
	    udiProfileVelocity := LREAL_TO_UDINT(ABS(Velocity) * Axis.fIncPerUnit));
	Done := _pp.xDone;
	Busy := _pp.xBusy;
	Active := _pp.xBusy;
	CommandAborted := FALSE;
	Error := _pp.xError;
	IF _pp.xError THEN ErrorID := SMC_MA_INVALID_ACCDEC_VALUES;
	ELSE ErrorID := SMC_NO_ERROR; END_IF
END_FUNCTION_BLOCK

(* ---------------------------------------------------------- MC_MoveRelative *)
FUNCTION_BLOCK MC_MoveRelative
VAR_IN_OUT
	Axis : AXIS_REF_SM3;
END_VAR
VAR_INPUT
	Execute : BOOL;
	Distance : LREAL;             (* [u] *)
	Velocity : LREAL;             (* [u/s] *)
	Acceleration : LREAL;
	Deceleration : LREAL;
	Jerk : LREAL;
	BufferMode : MC_BUFFER_MODE := mcbm_aborting;
END_VAR
VAR_OUTPUT
	Done : BOOL;
	Busy : BOOL;
	Active : BOOL;
	CommandAborted : BOOL;
	Error : BOOL;
	ErrorID : SMC_ERROR;
END_VAR
VAR
	_pp : OpenSML_ProfilePosition;
END_VAR
	IF Execute THEN
		Axis.byControllerMode := BYTE#3;
		Axis.fSetVelocity := Velocity;
	END_IF
	_pp(Axis := Axis.Drive,
	    xEnable := Execute,
	    xExecute := Execute,
	    xContinueMove := (BufferMode <> mcbm_aborting),
	    xRelativeMode := TRUE,
	    diTargetPosition := LREAL_TO_DINT(Distance * Axis.fIncPerUnit),
	    udiProfileVelocity := LREAL_TO_UDINT(ABS(Velocity) * Axis.fIncPerUnit));
	Done := _pp.xDone;
	Busy := _pp.xBusy;
	Active := _pp.xBusy;
	CommandAborted := FALSE;
	Error := _pp.xError;
	IF _pp.xError THEN ErrorID := SMC_MA_INVALID_ACCDEC_VALUES;
	ELSE ErrorID := SMC_NO_ERROR; END_IF
END_FUNCTION_BLOCK

(* ---------------------------------------------------------- MC_MoveVelocity *)
FUNCTION_BLOCK MC_MoveVelocity
VAR_IN_OUT
	Axis : AXIS_REF_SM3;
END_VAR
VAR_INPUT
	Execute : BOOL;
	Velocity : LREAL;             (* [u/s], signed *)
	Acceleration : LREAL;
	Deceleration : LREAL;
	Jerk : LREAL;
	Direction : MC_DIRECTION := mcd_current;
	BufferMode : MC_BUFFER_MODE := mcbm_aborting;
END_VAR
VAR_OUTPUT
	InVelocity : BOOL;
	Busy : BOOL;
	Active : BOOL;
	CommandAborted : BOOL;
	Error : BOOL;
	ErrorID : SMC_ERROR;
END_VAR
VAR
	_pv : OpenSML_ProfileVelocity;
END_VAR
	IF Execute THEN
		Axis.byControllerMode := BYTE#2;   (* SMC_velocity *)
		Axis.fSetVelocity := Velocity;
	END_IF
	_pv(Axis := Axis.Drive,
	    xEnable := Execute,
	    diTargetVelocity := LREAL_TO_DINT(Velocity * Axis.fIncPerUnit));
	Busy := Execute AND NOT _pv.xError;
	Active := Busy;
	CommandAborted := FALSE;
	Error := _pv.xError;
	(* target reached: commanded, no fault, and actual within 1% of target *)
	InVelocity := Execute AND NOT _pv.xError
	              AND (ABS(Axis.fActVelocity - Velocity) <= (ABS(Velocity) * 0.01 + 1.0));
	IF _pv.xError THEN ErrorID := SMC_MV_INVALID_VELACC_VALUES;
	ELSE ErrorID := SMC_NO_ERROR; END_IF
END_FUNCTION_BLOCK

(* ------------------------------------------------------------------- MC_Halt *)
FUNCTION_BLOCK MC_Halt
VAR_IN_OUT
	Axis : AXIS_REF_SM3;
END_VAR
VAR_INPUT
	Execute : BOOL;
	Deceleration : LREAL;
	Jerk : LREAL;
	BufferMode : MC_BUFFER_MODE := mcbm_aborting;
END_VAR
VAR_OUTPUT
	Done : BOOL;
	Busy : BOOL;
	Active : BOOL;
	CommandAborted : BOOL;
	Error : BOOL;
	ErrorID : SMC_ERROR;
END_VAR
VAR
	_stp : OpenSML_Stop;
END_VAR
	IF Execute THEN
		Axis.fSetDeceleration := Deceleration;
		Axis.fSetJerk := Jerk;
	END_IF
	_stp(Axis := Axis.Drive, xStop := Execute);
	(* standstill reached (SW bit14) => done; axis remains ready for new moves *)
	Done := Execute AND Axis.Drive.StatusWord.14;
	Busy := Execute AND NOT Done;
	Active := Busy;
	CommandAborted := FALSE;
	Error := Axis.Drive.StatusWord.3;
	IF Error THEN ErrorID := SMC_STOP_ERROR_DURING_STOP;
	ELSE ErrorID := SMC_NO_ERROR; END_IF
END_FUNCTION_BLOCK

(* ------------------------------------------------------------------- MC_Stop *)
FUNCTION_BLOCK MC_Stop
VAR_IN_OUT
	Axis : AXIS_REF_SM3;
END_VAR
VAR_INPUT
	Execute : BOOL;
	Deceleration : LREAL;
	Jerk : LREAL;
END_VAR
VAR_OUTPUT
	Done : BOOL;
	Busy : BOOL;
	Error : BOOL;
	ErrorID : SMC_ERROR;
END_VAR
VAR
	_stp : OpenSML_Stop;
END_VAR
	IF Execute THEN
		Axis.fSetDeceleration := Deceleration;
		Axis.fSetJerk := Jerk;
	END_IF
	(* MC_Stop locks the axis while Execute is held (no new motion accepted) *)
	_stp(Axis := Axis.Drive, xStop := Execute);
	Done := Execute AND Axis.Drive.StatusWord.14;
	Busy := Execute AND NOT Done;
	Error := Axis.Drive.StatusWord.3;
	IF Error THEN ErrorID := SMC_STOP_ERROR_DURING_STOP;
	ELSE ErrorID := SMC_NO_ERROR; END_IF
END_FUNCTION_BLOCK

(* ------------------------------------------------------------------ MC_Reset *)
FUNCTION_BLOCK MC_Reset
VAR_IN_OUT
	Axis : AXIS_REF_SM3;
END_VAR
VAR_INPUT
	Execute : BOOL;
END_VAR
VAR_OUTPUT
	Done : BOOL;
	Busy : BOOL;
	Error : BOOL;
	ErrorID : SMC_ERROR;
END_VAR
	(* CiA 402 fault reset (Controlword bit 7); Done when fault (SW bit3) clears *)
	Axis.Drive.ControlWord.7 := Execute;
	Done := Execute AND NOT Axis.Drive.StatusWord.3;
	Busy := Execute AND Axis.Drive.StatusWord.3;
	Error := FALSE;
	ErrorID := SMC_NO_ERROR;
END_FUNCTION_BLOCK

(* ------------------------------------------------------------------- MC_Home *)
FUNCTION_BLOCK MC_Home
VAR_IN_OUT
	Axis : AXIS_REF_SM3;
END_VAR
VAR_INPUT
	Execute : BOOL;
	Position : LREAL;             (* absolute position at reference [u] *)
END_VAR
VAR_OUTPUT
	Done : BOOL;
	Busy : BOOL;
	CommandAborted : BOOL;
	Error : BOOL;
	ErrorID : SMC_ERROR;
END_VAR
VAR
	_hm : OpenSML_Home;
END_VAR
	IF Execute THEN
		Axis.fSetPosition := Position;
	END_IF
	_hm(Axis := Axis.Drive, xEnable := Execute);
	Done := _hm.xDone;
	Busy := Execute AND NOT _hm.xDone AND NOT _hm.xError;
	CommandAborted := FALSE;
	Error := _hm.xError;
	IF _hm.xError THEN ErrorID := SMC_H_HOMING_TIMEOUT;
	ELSE ErrorID := SMC_NO_ERROR; END_IF
END_FUNCTION_BLOCK

(* ------------------------------------------------------------- MC_ReadStatus *)
FUNCTION_BLOCK MC_ReadStatus
VAR_IN_OUT
	Axis : AXIS_REF_SM3;
END_VAR
VAR_INPUT
	Enable : BOOL;
END_VAR
VAR_OUTPUT
	Valid : BOOL;
	Busy : BOOL;
	Error : BOOL;
	ErrorID : SMC_ERROR;
	Disabled : BOOL;
	Errorstop : BOOL;
	Stopping : BOOL;
	StandStill : BOOL;
	DiscreteMotion : BOOL;
	ContinuousMotion : BOOL;
	SynchronizedMotion : BOOL;
	Homing : BOOL;
	ConstantVelocity : BOOL;
	Accelerating : BOOL;
	Decelerating : BOOL;
	FBErrorOccured : BOOL;
END_VAR
	Valid := Enable;
	Busy := FALSE;
	IF Enable THEN
		Disabled := Axis.nAxisState = SMC_AXIS_STATE.power_off;
		Errorstop := Axis.nAxisState = SMC_AXIS_STATE.errorstop;
		Stopping := Axis.nAxisState = SMC_AXIS_STATE.stopping;
		StandStill := Axis.nAxisState = SMC_AXIS_STATE.standstill;
		DiscreteMotion := Axis.nAxisState = SMC_AXIS_STATE.discrete_motion;
		ContinuousMotion := Axis.nAxisState = SMC_AXIS_STATE.continuous_motion;
		SynchronizedMotion := Axis.nAxisState = SMC_AXIS_STATE.synchronized_motion;
		Homing := Axis.nAxisState = SMC_AXIS_STATE.homing;
		Error := Axis.bError;
		FBErrorOccured := Axis.bError;
		IF Axis.bError THEN ErrorID := SMC_DI_AXIS_ERROR;
		ELSE ErrorID := SMC_NO_ERROR; END_IF
	END_IF
END_FUNCTION_BLOCK

(* ------------------------------------------------------ MC_ReadActualPosition *)
FUNCTION_BLOCK MC_ReadActualPosition
VAR_IN_OUT
	Axis : AXIS_REF_SM3;
END_VAR
VAR_INPUT
	Enable : BOOL;
END_VAR
VAR_OUTPUT
	Valid : BOOL;
	Busy : BOOL;
	Error : BOOL;
	ErrorID : SMC_ERROR;
	Position : LREAL;             (* [u] *)
END_VAR
	Valid := Enable;
	Busy := FALSE;
	Error := FALSE;
	ErrorID := SMC_NO_ERROR;
	IF Enable THEN
		Position := Axis.fActPosition;
	END_IF
END_FUNCTION_BLOCK

(* ------------------------------------------------------ MC_ReadActualVelocity *)
FUNCTION_BLOCK MC_ReadActualVelocity
VAR_IN_OUT
	Axis : AXIS_REF_SM3;
END_VAR
VAR_INPUT
	Enable : BOOL;
END_VAR
VAR_OUTPUT
	Valid : BOOL;
	Busy : BOOL;
	Error : BOOL;
	ErrorID : SMC_ERROR;
	Velocity : LREAL;            (* [u/s] *)
END_VAR
	Valid := Enable;
	Busy := FALSE;
	Error := FALSE;
	ErrorID := SMC_NO_ERROR;
	IF Enable THEN
		Velocity := Axis.fActVelocity;
	END_IF
END_FUNCTION_BLOCK

(* ---------------------------------------------------------- MC_ReadAxisError *)
FUNCTION_BLOCK MC_ReadAxisError
VAR_IN_OUT
	Axis : AXIS_REF_SM3;
END_VAR
VAR_INPUT
	Enable : BOOL;
END_VAR
VAR_OUTPUT
	Valid : BOOL;
	Busy : BOOL;
	Error : BOOL;
	ErrorID : SMC_ERROR;
	AxisError : BOOL;
	AxisErrorID : DWORD;
END_VAR
	Valid := Enable;
	Busy := FALSE;
	Error := FALSE;
	ErrorID := SMC_NO_ERROR;
	IF Enable THEN
		AxisError := Axis.bError;
		AxisErrorID := Axis.dwErrorID;
	END_IF
END_FUNCTION_BLOCK
